      R_f[3,0] := -0.22841774;
      R_f[3,1] := 0.40559068;
      R_f[3,2] := 0.57486951;
      R_f[3,3] := 2.06207776;
      R_f[3,4] := -0.55732775;
      R_f[3,5] := 0.09659977;
      R_f[3,6] := -0.42354828;
      R_f[3,7] := -0.45963588;
      R_f[3,8] := -0.44553128;
      R_f[3,9] := -0.58046556;
      R_f[3,10] := -0.80908269;
      R_f[3,11] := -0.36142787;
      R_f[3,12] := 0.31985673;
      R_f[3,13] := -0.12466143;
      R_f[3,14] := 0.03553643;
      R_f[3,15] := -0.42549297;
      R_f[3,16] := -0.98859489;
      R_f[3,17] := 0.11508524;
      R_f[3,18] := 0.12030809;
      R_f[3,19] := 0.61023998;
      R_f[3,20] := -0.23926187;
      R_f[3,21] := -0.02740595;
      R_f[3,22] := 0.06562693;
      R_f[3,23] := 0.00750753;
      R_f[3,24] := 0.04459137;
      R_f[3,25] := 0.22271563;
      R_f[3,26] := -0.04020920;
      R_f[3,27] := 0.33254516;
      R_f[3,28] := 0.11126116;
      R_f[3,29] := -0.20861124;
      R_f[3,30] := 0.21898773;
      R_f[3,31] := 0.09003633;
      R_f[4,0] := -0.29503077;
      R_f[4,1] := 0.29277351;
      R_f[4,2] := -0.33615652;
      R_f[4,3] := 0.01891872;
      R_f[4,4] := -1.01232004;
      R_f[4,5] := 0.50957382;
      R_f[4,6] := -0.09908187;
      R_f[4,7] := -0.13480274;
      R_f[4,8] := -0.03347661;
      R_f[4,9] := 0.26127309;
      R_f[4,10] := -0.11804081;
      R_f[4,11] := -0.43345410;
      R_f[4,12] := 0.43429026;
      R_f[4,13] := -0.29253858;
      R_f[4,14] := 0.34731063;
      R_f[4,15] := -0.31193343;
      R_f[4,16] := 0.44109902;
      R_f[4,17] := 0.05499700;
      R_f[4,18] := -0.03124390;
      R_f[4,19] := -0.06733673;
      R_f[4,20] := 0.53314525;
      R_f[4,21] := 0.02740945;
      R_f[4,22] := -0.01510098;
      R_f[4,23] := 0.22094952;
      R_f[4,24] := -0.13394623;
      R_f[4,25] := 0.16025461;
      R_f[4,26] := 0.41375709;
      R_f[4,27] := -0.68666464;
      R_f[4,28] := 0.17169803;
      R_f[4,29] := -0.06553656;
      R_f[4,30] := -0.27536944;
      R_f[4,31] := 0.20692281;
      R_f[5,0] := 0.33732611;
      R_f[5,1] := 0.40928459;
      R_f[5,2] := -0.75300062;
      R_f[5,3] := -0.55881333;
      R_f[5,4] := 0.83829790;
      R_f[5,5] := -1.23661423;
      R_f[5,6] := -0.00860018;
      R_f[5,7] := 0.15366301;
      R_f[5,8] := 0.83814925;
      R_f[5,9] := -0.83846211;
      R_f[5,10] := 0.15663271;
      R_f[5,11] := -0.53920645;
      R_f[5,12] := -0.22816044;
      R_f[5,13] := -0.81048518;
      R_f[5,14] := 0.00169420;
      R_f[5,15] := 0.16230814;
      R_f[5,16] := 0.78781903;
      R_f[5,17] := -0.45289493;
      R_f[5,18] := 0.47988066;
      R_f[5,19] := -0.27889726;
      R_f[5,20] := 0.08924929;
      R_f[5,21] := -0.53515106;
      R_f[5,22] := 0.83308595;
      R_f[5,23] := 0.17609777;
      R_f[5,24] := -0.01040109;
      R_f[5,25] := 0.30510819;
      R_f[5,26] := 0.55807745;
      R_f[5,27] := 0.10998377;
      R_f[5,28] := -0.16242138;
      R_f[5,29] := -0.67912698;
      R_f[5,30] := -0.18073113;
      R_f[5,31] := 0.44595328;
      R_f[6,0] := -0.02960970;
      R_f[6,1] := 0.14120346;
      R_f[6,2] := -0.19232050;
      R_f[6,3] := -0.20220532;
      R_f[6,4] := 0.59759414;
      R_f[6,5] := 0.07536479;
      R_f[6,6] := 0.45140901;
      R_f[6,7] := -0.13872539;
      R_f[6,8] := 0.89296800;
      R_f[6,9] := -0.13736337;
      R_f[6,10] := 0.20182616;
      R_f[6,11] := -0.13915065;
      R_f[6,12] := -0.17636664;
      R_f[6,13] := -0.37117252;
      R_f[6,14] := 0.26237535;
      R_f[6,15] := -0.13584390;
      R_f[6,16] := 0.23492494;
      R_f[6,17] := -0.51170081;
      R_f[6,18] := -0.13849613;
      R_f[6,19] := -0.06773239;
      R_f[6,20] := 0.28203338;
      R_f[6,21] := 0.02628134;
      R_f[6,22] := 0.24086651;
      R_f[6,23] := 0.14421909;
      R_f[6,24] := 0.81928957;
      R_f[6,25] := 0.33552960;
      R_f[6,26] := -0.28975615;
      R_f[6,27] := 0.02547251;
      R_f[6,28] := 0.20271114;
      R_f[6,29] := -0.14385954;
      R_f[6,30] := 0.29766709;
      R_f[6,31] := -0.40624860;
      R_f[7,0] := 0.61828715;
      R_f[7,1] := 0.51957172;
      R_f[7,2] := 0.07738917;
      R_f[7,3] := -0.00875778;
      R_f[7,4] := 0.67404419;
      R_f[7,5] := 0.11073278;
      R_f[7,6] := -0.37006202;
      R_f[7,7] := 1.03556788;
      R_f[7,8] := 0.70712101;
      R_f[7,9] := -0.56803280;
      R_f[7,10] := -0.06974930;
      R_f[7,11] := 0.14248914;
      R_f[7,12] := 0.66664493;
      R_f[7,13] := -0.50647444;
      R_f[7,14] := 0.28662270;
      R_f[7,15] := 0.16329370;
      R_f[7,16] := -0.00441234;
      R_f[7,17] := -0.22685143;
      R_f[7,18] := -0.64886677;
      R_f[7,19] := -0.03913877;
      R_f[7,20] := 0.57906586;
      R_f[7,21] := 0.41091961;
      R_f[7,22] := 0.19402935;
      R_f[7,23] := -0.56783932;
      R_f[7,24] := 0.59809852;
      R_f[7,25] := 0.22131553;
      R_f[7,26] := 0.01115896;
      R_f[7,27] := 0.20468640;
      R_f[7,28] := -0.69074368;
      R_f[7,29] := -0.22870129;
      R_f[7,30] := 0.38742521;
      R_f[7,31] := -0.17464639;
      R_f[8,0] := -0.01413119;
      R_f[8,1] := -0.01563436;
      R_f[8,2] := 0.04907341;
      R_f[8,3] := 0.13082743;
      R_f[8,4] := -0.14134008;
      R_f[8,5] := -0.09485538;
      R_f[8,6] := -0.31782639;
      R_f[8,7] := -0.00754579;
      R_f[8,8] := -0.68271863;
      R_f[8,9] := 0.43590066;
      R_f[8,10] := -0.16523221;
      R_f[8,11] := 0.20073125;
      R_f[8,12] := -0.47652704;
      R_f[8,13] := 0.18128465;
      R_f[8,14] := -0.62839359;
      R_f[8,15] := -0.25646719;
      R_f[8,16] := -0.23885600;
      R_f[8,17] := 0.13142671;
      R_f[8,18] := 0.48771819;
      R_f[8,19] := -0.49085858;
      R_f[8,20] := -0.18839863;
      R_f[8,21] := -0.43685639;
      R_f[8,22] := 0.02705371;
      R_f[8,23] := -0.05543226;
      R_f[8,24] := -0.38585073;
      R_f[8,25] := 0.06531966;
      R_f[8,26] := -0.15446883;
      R_f[8,27] := 0.05854914;
      R_f[8,28] := -0.30904549;
      R_f[8,29] := 0.05056802;
      R_f[8,30] := -0.41357008;
      R_f[8,31] := 0.20621774;
      R_f[9,0] := -0.83740795;
      R_f[9,1] := -0.06988145;
      R_f[9,2] := -0.01356161;
      R_f[9,3] := 0.08127308;
      R_f[9,4] := -0.45402661;
      R_f[9,5] := 0.38458407;
      R_f[9,6] := 0.26937473;
      R_f[9,7] := -0.32646099;
      R_f[9,8] := -0.91716331;
      R_f[9,9] := 1.38183928;
      R_f[9,10] := 0.15634774;
      R_f[9,11] := -0.17276365;
      R_f[9,12] := -0.16843350;
      R_f[9,13] := -0.24043344;
      R_f[9,14] := -1.08728600;
      R_f[9,15] := -0.43865058;
      R_f[9,16] := 0.03624129;
      R_f[9,17] := 0.46195465;
      R_f[9,18] := 0.28181869;
      R_f[9,19] := 0.00515404;
      R_f[9,20] := -0.05451173;
      R_f[9,21] := 0.29636249;
      R_f[9,22] := -0.61817378;
      R_f[9,23] := 0.29860359;
      R_f[9,24] := -0.34871268;
      R_f[9,25] := 0.11697577;
      R_f[9,26] := 0.78417259;
      R_f[9,27] := 0.71926928;
      R_f[9,28] := -0.20325977;
      R_f[9,29] := 0.14632353;
      R_f[9,30] := -0.25228071;
      R_f[9,31] := -0.32943490;
      R_f[10,0] := 0.38591698;
      R_f[10,1] := 0.00522286;
      R_f[10,2] := -0.48348549;
      R_f[10,3] := 0.96521038;
      R_f[10,4] := -0.32313466;
      R_f[10,5] := 0.30804583;
      R_f[10,6] := -0.79955953;
      R_f[10,7] := -0.31883714;
      R_f[10,8] := -0.90835553;
      R_f[10,9] := 0.30884159;
      R_f[10,10] := -1.16350293;
      R_f[10,11] := -0.63253200;
      R_f[10,12] := 0.59796506;
      R_f[10,13] := 0.48238036;
      R_f[10,14] := -0.10394208;
      R_f[10,15] := 0.16137904;
      R_f[10,16] := 0.11384938;
      R_f[10,17] := 1.00142598;
      R_f[10,18] := -0.75928485;
      R_f[10,19] := 0.28338146;
      R_f[10,20] := -0.95777762;
      R_f[10,21] := -0.61350137;
      R_f[10,22] := -0.70301116;
      R_f[10,23] := 0.22109440;
      R_f[10,24] := 0.32511491;
      R_f[10,25] := 0.58860904;
      R_f[10,26] := -0.02545941;
      R_f[10,27] := 0.26207218;
      R_f[10,28] := 0.75892609;
      R_f[10,29] := -0.47240314;
      R_f[10,30] := 0.02046607;
      R_f[10,31] := -0.29343525;
      R_f[11,0] := 0.63524234;
      R_f[11,1] := 0.13768600;
      R_f[11,2] := -0.28915507;
      R_f[11,3] := -0.18023908;
      R_f[11,4] := -0.26212382;
      R_f[11,5] := -0.55292249;
      R_f[11,6] := 0.16202901;
      R_f[11,7] := 0.35055608;
      R_f[11,8] := 0.59746683;
      R_f[11,9] := -0.60563761;
      R_f[11,10] := -0.04891396;
      R_f[11,11] := 1.17771423;
      R_f[11,12] := -0.31640816;
      R_f[11,13] := -0.11039021;
      R_f[11,14] := -0.08756445;
      R_f[11,15] := 0.00601315;
      R_f[11,16] := 0.32191852;
      R_f[11,17] := -0.90107346;
      R_f[11,18] := -0.47469705;
      R_f[11,19] := 0.05416169;
      R_f[11,20] := -0.09831773;
      R_f[11,21] := 0.10362659;
      R_f[11,22] := -0.00615723;
      R_f[11,23] := -0.13419445;
      R_f[11,24] := 0.07473942;
      R_f[11,25] := 0.45523170;
      R_f[11,26] := 0.17231539;
      R_f[11,27] := 0.18330109;
      R_f[11,28] := -0.33154044;
      R_f[11,29] := 0.00715767;
      R_f[11,30] := 0.02798121;
      R_f[11,31] := 0.12936890;
      R_f[12,0] := 0.52463913;
      R_f[12,1] := 1.23480833;
      R_f[12,2] := -0.26183358;
      R_f[12,3] := 0.29687256;
      R_f[12,4] := 0.12944640;
      R_f[12,5] := -0.64208639;
      R_f[12,6] := 0.14092363;
      R_f[12,7] := 0.29900426;
      R_f[12,8] := -0.38989353;
      R_f[12,9] := -0.15832269;
      R_f[12,10] := 0.38569406;
      R_f[12,11] := -0.49528036;
      R_f[12,12] := 0.83373916;
      R_f[12,13] := -0.42694458;
      R_f[12,14] := 0.76566309;
      R_f[12,15] := -0.48013216;
      R_f[12,16] := 0.40656197;
      R_f[12,17] := -0.31445476;
      R_f[12,18] := 0.24111255;
      R_f[12,19] := -0.19961938;
      R_f[12,20] := -0.11154682;
      R_f[12,21] := 0.33029765;
      R_f[12,22] := -0.13147451;
      R_f[12,23] := -0.03679356;
      R_f[12,24] := 0.17805246;
      R_f[12,25] := 0.05382822;
      R_f[12,26] := 0.43463483;
      R_f[12,27] := 0.27920336;
      R_f[12,28] := 0.55672109;
      R_f[12,29] := -0.69647855;
      R_f[12,30] := 0.65581310;
      R_f[12,31] := 0.12511645;
      R_f[13,0] := 0.23202457;
      R_f[13,1] := 0.62695414;
      R_f[13,2] := -0.71075511;
      R_f[13,3] := -0.91361868;
      R_f[13,4] := 1.39223123;
      R_f[13,5] := 0.40526325;
      R_f[13,6] := 0.07239435;
      R_f[13,7] := 0.16743791;
      R_f[13,8] := 0.89612418;
      R_f[13,9] := -0.92080438;
      R_f[13,10] := 0.23565021;
      R_f[13,11] := 0.41098762;
      R_f[13,12] := -0.37411463;
      R_f[13,13] := -0.37083071;
      R_f[13,14] := 0.21330817;
      R_f[13,15] := 0.32418102;
      R_f[13,16] := 0.64384466;
      R_f[13,17] := -0.70755357;
      R_f[13,18] := -0.60732776;
      R_f[13,19] := -0.31852406;
      R_f[13,20] := 0.38003522;
      R_f[13,21] := -0.38526192;
      R_f[13,22] := 0.85999751;
      R_f[13,23] := 0.08276569;
      R_f[13,24] := 0.52139038;
      R_f[13,25] := -0.09750945;
      R_f[13,26] := -0.19196609;
      R_f[13,27] := -0.18892166;
      R_f[13,28] := 0.12520945;
      R_f[13,29] := -0.40455785;
      R_f[13,30] := 0.87176305;
      R_f[13,31] := -0.29801390;
      R_f[14,0] := 0.08073674;
      R_f[14,1] := -0.22958316;
      R_f[14,2] := 0.39506468;
      R_f[14,3] := -0.29865783;
      R_f[14,4] := -0.24071212;
      R_f[14,5] := -0.54502225;
      R_f[14,6] := -0.22081053;
      R_f[14,7] := 0.11199540;
      R_f[14,8] := 0.39893955;
      R_f[14,9] := -0.00592328;
      R_f[14,10] := -0.56832987;
      R_f[14,11] := 0.19659449;
      R_f[14,12] := 0.57248878;
      R_f[14,13] := 0.22812998;
      R_f[14,14] := -0.08929932;
      R_f[14,15] := -0.43194354;
      R_f[14,16] := 0.15896702;
      R_f[14,17] := -0.12431962;
      R_f[14,18] := 0.43860698;
      R_f[14,19] := -0.23576687;
      R_f[14,20] := 0.12837251;
      R_f[14,21] := -0.08831814;
      R_f[14,22] := -0.12136080;
      R_f[14,23] := 0.56518930;
      R_f[14,24] := -0.46596053;
      R_f[14,25] := 0.19473872;
      R_f[14,26] := 0.19937690;
      R_f[14,27] := -1.21616924;
      R_f[14,28] := 0.46861416;
      R_f[14,29] := -0.24986319;
      R_f[14,30] := -0.61549062;
      R_f[14,31] := 0.33290240;
      R_f[15,0] := 0.31359208;
      R_f[15,1] := 0.33051741;
      R_f[15,2] := 0.15030840;
      R_f[15,3] := -0.38865900;
      R_f[15,4] := 0.06516448;
      R_f[15,5] := -0.32763284;
      R_f[15,6] := 0.21778707;
      R_f[15,7] := 0.23249651;
      R_f[15,8] := 0.02938646;
      R_f[15,9] := 0.06135718;
      R_f[15,10] := -0.27028698;
      R_f[15,11] := 0.40001541;
      R_f[15,12] := -0.00793086;
      R_f[15,13] := 0.00380884;
      R_f[15,14] := 0.08370329;
      R_f[15,15] := -0.22548552;
      R_f[15,16] := 0.02933858;
      R_f[15,17] := -0.35302344;
      R_f[15,18] := -0.25063863;
      R_f[15,19] := 0.28370765;
      R_f[15,20] := 0.04397562;
      R_f[15,21] := -0.07230925;
      R_f[15,22] := -0.09505362;
      R_f[15,23] := 0.15444055;
      R_f[15,24] := -0.02045420;
      R_f[15,25] := -0.14273162;
      R_f[15,26] := 0.37428376;
      R_f[15,27] := -0.05992498;
      R_f[15,28] := 0.16830987;
      R_f[15,29] := -0.32088986;
      R_f[15,30] := -0.33436120;
      R_f[15,31] := -0.37953538;
      R_f[16,0] := -0.26587957;
      R_f[16,1] := -0.31207001;
      R_f[16,2] := 0.50653142;
      R_f[16,3] := 1.14224505;
      R_f[16,4] := -0.61703724;
      R_f[16,5] := 0.13980502;
      R_f[16,6] := -0.14207593;
      R_f[16,7] := 0.39799580;
      R_f[16,8] := -0.42795599;
      R_f[16,9] := 0.49218190;
      R_f[16,10] := -0.02379325;
      R_f[16,11] := -0.01251386;
      R_f[16,12] := 0.81707931;
      R_f[16,13] := 0.56178325;
      R_f[16,14] := -0.41181156;
      R_f[16,15] := -0.34066352;
      R_f[16,16] := -0.47481647;
      R_f[16,17] := 0.51806176;
      R_f[16,18] := 0.20107090;
      R_f[16,19] := 0.04892090;
      R_f[16,20] := -0.22273828;
      R_f[16,21] := 0.42268997;
      R_f[16,22] := -0.21690965;
      R_f[16,23] := 0.55266404;
      R_f[16,24] := -0.78800714;
      R_f[16,25] := -0.40029246;
      R_f[16,26] := 0.31856278;
      R_f[16,27] := 0.15422256;
      R_f[16,28] := 0.08612204;
      R_f[16,29] := 0.27195919;
      R_f[16,30] := -0.04387485;
      R_f[16,31] := -0.06196566;
      R_f[17,0] := 0.05910539;
      R_f[17,1] := -0.21845020;
      R_f[17,2] := -0.64325720;
      R_f[17,3] := -0.17311564;
      R_f[17,4] := -0.05836086;
      R_f[17,5] := 0.08543847;
      R_f[17,6] := 0.43946153;
      R_f[17,7] := 0.30724356;
      R_f[17,8] := 0.06860433;
      R_f[17,9] := 0.62805259;
      R_f[17,10] := 0.54351902;
      R_f[17,11] := 0.07233211;
      R_f[17,12] := -0.29924318;
      R_f[17,13] := -0.46094373;
      R_f[17,14] := -0.06874729;
      R_f[17,15] := 0.24842280;
      R_f[17,16] := -0.51377529;
      R_f[17,17] := 1.53367448;
      R_f[17,18] := 0.33991754;
      R_f[17,19] := 0.21408086;
      R_f[17,20] := -0.02237522;
      R_f[17,21] := -0.02311720;
      R_f[17,22] := 0.23792864;
      R_f[17,23] := 0.21117508;
      R_f[17,24] := -0.01755552;
      R_f[17,25] := -0.14541535;
      R_f[17,26] := 0.62708884;
      R_f[17,27] := 0.03084901;
      R_f[17,28] := -0.38820636;
      R_f[17,29] := -0.19554625;
      R_f[17,30] := 0.06806003;
      R_f[17,31] := -0.30774286;
      R_f[18,0] := 0.16866495;
      R_f[18,1] := 0.42400992;
      R_f[18,2] := -0.36475778;
      R_f[18,3] := -0.46353397;
      R_f[18,4] := -0.23605427;
      R_f[18,5] := -0.39058918;
      R_f[18,6] := 0.24388304;
      R_f[18,7] := -0.24780002;
      R_f[18,8] := -0.12100184;
      R_f[18,9] := -0.35586256;
      R_f[18,10] := 0.54968441;
      R_f[18,11] := -0.25823474;
      R_f[18,12] := -0.37975135;
      R_f[18,13] := 0.10739443;
      R_f[18,14] := 0.02995439;
      R_f[18,15] := 0.37767676;
      R_f[18,16] := -0.06366078;
      R_f[18,17] := 0.32446918;
      R_f[18,18] := 0.87205279;
      R_f[18,19] := -0.05647478;
      R_f[18,20] := -0.19952400;
      R_f[18,21] := -0.61423117;
      R_f[18,22] := 0.49618649;
      R_f[18,23] := -0.15967572;
      R_f[18,24] := 0.65420824;
      R_f[18,25] := 0.12151071;
      R_f[18,26] := 0.31860438;
      R_f[18,27] := 0.02739185;
      R_f[18,28] := -0.66384917;
      R_f[18,29] := 0.17025499;
      R_f[18,30] := -0.25605354;
      R_f[18,31] := 0.52890509;
      R_f[19,0] := 0.65365380;
      R_f[19,1] := 0.10235491;
      R_f[19,2] := 0.62065804;
      R_f[19,3] := 0.10225008;
      R_f[19,4] := -0.45779619;
      R_f[19,5] := -0.42509148;
      R_f[19,6] := -0.48240736;
      R_f[19,7] := -0.41890648;
      R_f[19,8] := 0.51948655;
      R_f[19,9] := 0.22051780;
      R_f[19,10] := -0.32477748;
      R_f[19,11] := -1.20024562;
      R_f[19,12] := 0.22928596;
      R_f[19,13] := 0.10820945;
      R_f[19,14] := -0.23491700;
      R_f[19,15] := -0.34898815;
      R_f[19,16] := -0.93565780;
      R_f[19,17] := 0.20988458;
      R_f[19,18] := -0.31584072;
      R_f[19,19] := -0.02921623;
      R_f[19,20] := -0.26133105;
      R_f[19,21] := 0.63414830;
      R_f[19,22] := -0.26187015;
      R_f[19,23] := 0.26986319;
      R_f[19,24] := -0.16388878;
      R_f[19,25] := 0.39682811;
      R_f[19,26] := 0.23186836;
      R_f[19,27] := 0.33898479;
      R_f[19,28] := -0.19298120;
      R_f[19,29] := 0.05988296;
      R_f[19,30] := 0.30527696;
      R_f[19,31] := 0.35504943;
      R_f[20,0] := 0.60740626;
      R_f[20,1] := 0.68342733;
      R_f[20,2] := -0.56973433;
      R_f[20,3] := 0.30702043;
      R_f[20,4] := 0.63084090;
      R_f[20,5] := -0.76327389;
      R_f[20,6] := -0.16775738;
      R_f[20,7] := 0.29119602;
      R_f[20,8] := -0.24701932;
      R_f[20,9] := -0.93371648;
      R_f[20,10] := 0.65781426;
      R_f[20,11] := -0.03017730;
      R_f[20,12] := -0.59253180;
      R_f[20,13] := -1.06371450;
      R_f[20,14] := 0.88938069;
      R_f[20,15] := 0.20159939;
      R_f[20,16] := 0.31710625;
      R_f[20,17] := 0.17246717;
      R_f[20,18] := 0.76323175;
      R_f[20,19] := 0.10229112;
      R_f[20,20] := -0.21142122;
      R_f[20,21] := -0.31407952;
      R_f[20,22] := -0.34694698;
      R_f[20,23] := -0.14305308;
      R_f[20,24] := 0.66643405;
      R_f[20,25] := -0.32228628;
      R_f[20,26] := 0.18264067;
      R_f[20,27] := 0.21311571;
      R_f[20,28] := 0.15977044;
      R_f[20,29] := 0.35266665;
      R_f[20,30] := 0.07271075;
      R_f[20,31] := 0.90672767;
      R_f[21,0] := 0.63794458;
      R_f[21,1] := -0.07306197;
      R_f[21,2] := -0.33461115;
      R_f[21,3] := 0.07822674;
      R_f[21,4] := 0.38671464;
      R_f[21,5] := -0.92790735;
      R_f[21,6] := -0.12789188;
      R_f[21,7] := -0.12363939;
      R_f[21,8] := 0.18649052;
      R_f[21,9] := -0.47208816;
      R_f[21,10] := -0.51584691;
      R_f[21,11] := 0.18042590;
      R_f[21,12] := 0.45089826;
      R_f[21,13] := 0.13358073;
      R_f[21,14] := 0.68462294;
      R_f[21,15] := -0.50330412;
      R_f[21,16] := -0.00928727;
      R_f[21,17] := -0.18551630;
      R_f[21,18] := 0.23045629;
      R_f[21,19] := -0.24903311;
      R_f[21,20] := -0.21607880;
      R_f[21,21] := 1.09473407;
      R_f[21,22] := 0.22049566;
      R_f[21,23] := 0.00980196;
      R_f[21,24] := 0.42017451;
      R_f[21,25] := 0.18463401;
      R_f[21,26] := 0.72073048;
      R_f[21,27] := 0.08499105;
      R_f[21,28] := -0.05317052;
      R_f[21,29] := 0.01483204;
      R_f[21,30] := 0.42573896;
      R_f[21,31] := 0.58880693;
      R_f[22,0] := 0.52571583;
      R_f[22,1] := 0.74352360;
      R_f[22,2] := -0.42845920;
      R_f[22,3] := -0.12134498;
      R_f[22,4] := -0.33517385;
      R_f[22,5] := -0.53988433;
      R_f[22,6] := -0.19025023;
      R_f[22,7] := -0.33218449;
      R_f[22,8] := -0.56198525;
      R_f[22,9] := 0.06062734;
      R_f[22,10] := -0.15277702;
      R_f[22,11] := -0.15610690;
      R_f[22,12] := -0.85074830;
      R_f[22,13] := -0.27995047;
      R_f[22,14] := 0.04608161;
      R_f[22,15] := 0.20265953;
      R_f[22,16] := 0.61842918;
      R_f[22,17] := -0.35963365;
      R_f[22,18] := 0.32028535;
      R_f[22,19] := 0.40971312;
      R_f[22,20] := 0.07105415;
      R_f[22,21] := -0.26550075;
      R_f[22,22] := 0.32755789;
      R_f[22,23] := -0.53670889;
      R_f[22,24] := 0.81352252;
      R_f[22,25] := 0.17814557;
      R_f[22,26] := -0.27500603;
      R_f[22,27] := 0.17979041;
      R_f[22,28] := 0.77811944;
      R_f[22,29] := -0.40859875;
      R_f[22,30] := -0.01199397;
      R_f[22,31] := 0.16662607;
      R_f[23,0] := 0.18513951;
      R_f[23,1] := -0.36498722;
      R_f[23,2] := 0.12142582;
      R_f[23,3] := 0.06119955;
      R_f[23,4] := 0.18143424;
      R_f[23,5] := -0.15825206;
      R_f[23,6] := -0.56776536;
      R_f[23,7] := 0.03979553;
      R_f[23,8] := -0.57782358;
      R_f[23,9] := 0.17007102;
      R_f[23,10] := 0.03401264;
      R_f[23,11] := 0.30232838;
      R_f[23,12] := 0.60225219;
      R_f[23,13] := 0.13679615;
      R_f[23,14] := -0.17490226;
      R_f[23,15] := -0.38221130;
      R_f[23,16] := -0.35548767;
      R_f[23,17] := -0.11720476;
      R_f[23,18] := 0.10709175;
      R_f[23,19] := 0.27031457;
      R_f[23,20] := -0.21203364;
      R_f[23,21] := 0.10817976;
      R_f[23,22] := -0.02741619;
      R_f[23,23] := -0.12317895;
      R_f[23,24] := -0.43592772;
      R_f[23,25] := -0.06452787;
      R_f[23,26] := 0.23145935;
      R_f[23,27] := -0.13228178;
      R_f[23,28] := -0.27505627;
      R_f[23,29] := 0.07636941;
      R_f[23,30] := -0.40810692;
      R_f[23,31] := 0.42898092;
      R_f[24,0] := 0.28041553;
      R_f[24,1] := 0.35192281;
      R_f[24,2] := -0.45653370;
      R_f[24,3] := -0.39068758;
      R_f[24,4] := 0.59820068;
      R_f[24,5] := -0.14331487;
      R_f[24,6] := -0.16312519;
      R_f[24,7] := 0.20082375;
      R_f[24,8] := 0.85522902;
      R_f[24,9] := -1.29532707;
      R_f[24,10] := 0.44740444;
      R_f[24,11] := -0.42685062;
      R_f[24,12] := -0.38446230;
      R_f[24,13] := -0.25391304;
      R_f[24,14] := 0.57489002;
      R_f[24,15] := -0.11480054;
      R_f[24,16] := 0.49371004;
      R_f[24,17] := -0.34504244;
      R_f[24,18] := 0.08720941;
      R_f[24,19] := -0.72877926;
      R_f[24,20] := -0.04864010;
      R_f[24,21] := -0.53587073;
      R_f[24,22] := 0.82679683;
      R_f[24,23] := -0.64950413;
      R_f[24,24] := 0.71601194;
      R_f[24,25] := 0.38295448;
      R_f[24,26] := 0.40242442;
      R_f[24,27] := 0.20521010;
      R_f[24,28] := -0.03906753;
      R_f[24,29] := -0.60810322;
      R_f[24,30] := 0.03209632;
      R_f[24,31] := -0.01952329;
      R_f[25,0] := 0.24457985;
      R_f[25,1] := -1.02144086;
      R_f[25,2] := -1.15114701;
      R_f[25,3] := -0.35912865;
      R_f[25,4] := 0.10526828;
      R_f[25,5] := -0.20179662;
      R_f[25,6] := -0.08682156;
      R_f[25,7] := -0.53071922;
      R_f[25,8] := 0.78854895;
      R_f[25,9] := -0.39259291;
      R_f[25,10] := 0.01843655;
      R_f[25,11] := -0.56601465;
      R_f[25,12] := -0.02357278;
      R_f[25,13] := -0.37074372;
      R_f[25,14] := -0.04764435;
      R_f[25,15] := 0.07631879;
      R_f[25,16] := 0.14908385;
      R_f[25,17] := -0.22848843;
      R_f[25,18] := 0.07038445;
      R_f[25,19] := -0.21256164;
      R_f[25,20] := -0.51917696;
      R_f[25,21] := -0.13761941;
      R_f[25,22] := 1.10180664;
      R_f[25,23] := -0.01601213;
      R_f[25,24] := 0.33799487;
      R_f[25,25] := 0.74898493;
      R_f[25,26] := 0.10358041;
      R_f[25,27] := -0.17927809;
      R_f[25,28] := -0.14816135;
      R_f[25,29] := -0.15051788;
      R_f[25,30] := 0.32431662;
      R_f[25,31] := -0.06228854;
      R_f[26,0] := -0.17391884;
      R_f[26,1] := 0.40459314;
      R_f[26,2] := 0.23582034;
      R_f[26,3] := 0.27855241;
      R_f[26,4] := 0.41587636;
      R_f[26,5] := -0.06871118;
      R_f[26,6] := -0.18198022;
      R_f[26,7] := 0.30424389;
      R_f[26,8] := 0.47402722;
      R_f[26,9] := 0.10770813;
      R_f[26,10] := 0.19400623;
      R_f[26,11] := 0.19763534;
      R_f[26,12] := 0.83919579;
      R_f[26,13] := -0.20429327;
      R_f[26,14] := 0.30284089;
      R_f[26,15] := -0.15002888;
      R_f[26,16] := 0.68186575;
      R_f[26,17] := 0.55425143;
      R_f[26,18] := 0.27912667;
      R_f[26,19] := 0.33006024;
      R_f[26,20] := 0.64902514;
      R_f[26,21] := -0.04681511;
      R_f[26,22] := 0.43274990;
      R_f[26,23] := -0.06403653;
      R_f[26,24] := 0.90166181;
      R_f[26,25] := -0.52762878;
      R_f[26,26] := -0.00969170;
      R_f[26,27] := -0.59007823;
      R_f[26,28] := 0.04513381;
      R_f[26,29] := -1.11053836;
      R_f[26,30] := -0.14078638;
      R_f[26,31] := 0.10301355;
      R_f[27,0] := 0.39776009;
      R_f[27,1] := 0.59193295;
      R_f[27,2] := -0.16674590;
      R_f[27,3] := -0.01398129;
      R_f[27,4] := 0.34197676;
      R_f[27,5] := -0.11277734;
      R_f[27,6] := -0.18087836;
      R_f[27,7] := -0.24809147;
      R_f[27,8] := 1.11544597;
      R_f[27,9] := -0.41635385;
      R_f[27,10] := 1.21610570;
      R_f[27,11] := -0.42330170;
      R_f[27,12] := -0.49244744;
      R_f[27,13] := -0.17151001;
      R_f[27,14] := -0.73654294;
      R_f[27,15] := 0.40863410;
      R_f[27,16] := 0.30207148;
      R_f[27,17] := -0.30706853;
      R_f[27,18] := 0.17934655;
      R_f[27,19] := -0.01947166;
      R_f[27,20] := 0.29237783;
      R_f[27,21] := -0.18835185;
      R_f[27,22] := -0.42462611;
      R_f[27,23] := -0.31352675;
      R_f[27,24] := 0.80565614;
      R_f[27,25] := 0.15593880;
      R_f[27,26] := -0.07164915;
      R_f[27,27] := 1.59558272;
      R_f[27,28] := -0.26499027;
      R_f[27,29] := -0.86730254;
      R_f[27,30] := 0.45258304;
      R_f[27,31] := -0.10650399;
      R_f[28,0] := 0.29013574;
      R_f[28,1] := 0.78875935;
      R_f[28,2] := -0.22047451;
      R_f[28,3] := 0.31630492;
      R_f[28,4] := 0.13784394;
      R_f[28,5] := -0.17747335;
      R_f[28,6] := -0.16462083;
      R_f[28,7] := 0.02444983;
      R_f[28,8] := 0.02157918;
      R_f[28,9] := -0.85899609;
      R_f[28,10] := 0.51003945;
      R_f[28,11] := 0.22153500;
      R_f[28,12] := -0.81957668;
      R_f[28,13] := 0.15229519;
      R_f[28,14] := -0.49981925;
      R_f[28,15] := -0.20841819;
      R_f[28,16] := 0.48134491;
      R_f[28,17] := -0.58209991;
      R_f[28,18] := -0.21895251;
      R_f[28,19] := -0.31777707;
      R_f[28,20] := 0.39952904;
      R_f[28,21] := 0.33487400;
      R_f[28,22] := 0.53231794;
      R_f[28,23] := 0.58753723;
      R_f[28,24] := 0.29652479;
      R_f[28,25] := 0.49816924;
      R_f[28,26] := -0.19129919;
      R_f[28,27] := 0.74723542;
      R_f[28,28] := 0.06283404;
      R_f[28,29] := -0.70639998;
      R_f[28,30] := 0.34521261;
      R_f[28,31] := -0.15957113;
      R_f[29,0] := 0.23835732;
      R_f[29,1] := -0.26068553;
      R_f[29,2] := -0.55099136;
      R_f[29,3] := -0.27018866;
      R_f[29,4] := -0.35758555;
      R_f[29,5] := 0.74466068;
      R_f[29,6] := 0.46339175;
      R_f[29,7] := -0.27842417;
      R_f[29,8] := 0.12199467;
      R_f[29,9] := -0.58916980;
      R_f[29,10] := 0.10298276;
      R_f[29,11] := -0.58598566;
      R_f[29,12] := 0.03986860;
      R_f[29,13] := 0.36140522;
      R_f[29,14] := 0.14722234;
      R_f[29,15] := -0.15363480;
      R_f[29,16] := 0.72394967;
      R_f[29,17] := -0.39522561;
      R_f[29,18] := -0.06369760;
      R_f[29,19] := -0.19733445;
      R_f[29,20] := -0.23108549;
      R_f[29,21] := 0.09581164;
      R_f[29,22] := 0.60348934;
      R_f[29,23] := 0.38583145;
      R_f[29,24] := -0.32982609;
      R_f[29,25] := 0.76995927;
      R_f[29,26] := 0.39173558;
      R_f[29,27] := -0.11436092;
      R_f[29,28] := -0.33975780;
      R_f[29,29] := -2.43963838;
      R_f[29,30] := 0.01613091;
      R_f[29,31] := 1.01884580;
      R_f[30,0] := 0.44902706;
      R_f[30,1] := -0.01531547;
      R_f[30,2] := 0.43428138;
      R_f[30,3] := 0.20990226;
      R_f[30,4] := 0.10665958;
      R_f[30,5] := -0.07787514;
      R_f[30,6] := -0.28534907;
      R_f[30,7] := -0.20589265;
      R_f[30,8] := -0.26249862;
      R_f[30,9] := 0.32755303;
      R_f[30,10] := 0.16526289;
      R_f[30,11] := 0.07607982;
      R_f[30,12] := 0.15522026;
      R_f[30,13] := 0.16349413;
      R_f[30,14] := -0.41222379;
      R_f[30,15] := -0.37317255;
      R_f[30,16] := -0.38004446;
      R_f[30,17] := -0.11156923;
      R_f[30,18] := -0.06939796;
      R_f[30,19] := 0.75725025;
      R_f[30,20] := 0.16113472;
      R_f[30,21] := 0.36386901;
      R_f[30,22] := 0.15552250;
      R_f[30,23] := -0.10594840;
      R_f[30,24] := -0.00384362;
      R_f[30,25] := -0.10023083;
      R_f[30,26] := 0.55560988;
      R_f[30,27] := 0.35110676;
      R_f[30,28] := -0.28105840;
      R_f[30,29] := -0.08273152;
      R_f[30,30] := 0.76468736;
      R_f[30,31] := 0.03726526;
      R_f[31,0] := 0.43319872;
      R_f[31,1] := 0.89265436;
      R_f[31,2] := -0.02175743;
      R_f[31,3] := -0.23646763;
      R_f[31,4] := -0.24073155;
      R_f[31,5] := -0.00261918;
      R_f[31,6] := -0.57301140;
      R_f[31,7] := -0.04121628;
      R_f[31,8] := -0.32528654;
      R_f[31,9] := -0.79124427;
      R_f[31,10] := -0.25563994;
      R_f[31,11] := 0.61876816;
      R_f[31,12] := -0.24966605;
      R_f[31,13] := -0.15887363;
      R_f[31,14] := -0.27610224;
      R_f[31,15] := -0.24292535;
      R_f[31,16] := -0.17999788;
      R_f[31,17] := -0.17289916;
      R_f[31,18] := 0.49396884;
      R_f[31,19] := 0.35957804;
      R_f[31,20] := -0.07121407;
      R_f[31,21] := 0.01738700;
      R_f[31,22] := 0.34174326;
      R_f[31,23] := -0.52943313;
      R_f[31,24] := -0.28900346;
      R_f[31,25] := 0.48076582;
      R_f[31,26] := -0.03657150;
      R_f[31,27] := 0.02927713;
      R_f[31,28] := -0.82611400;
      R_f[31,29] := -0.81384391;
      R_f[31,30] := -0.24894159;
      R_f[31,31] := 1.24944818;
      R_g[0,0] := -3.90892291;
      R_g[0,1] := -0.07594703;
      R_g[0,2] := -0.11032616;
      R_g[0,3] := -0.12472310;
      R_g[0,4] := -0.00621575;
      R_g[0,5] := 0.19935456;
      R_g[0,6] := -0.06362464;
      R_g[0,7] := -0.16034737;
      R_g[0,8] := 0.09810749;
      R_g[0,9] := 0.12010512;
      R_g[0,10] := 0.17773002;
      R_g[0,11] := -0.01798855;
      R_g[0,12] := -0.10235326;
      R_g[0,13] := 0.23832326;
      R_g[0,14] := 0.11828293;
      R_g[0,15] := -0.07939270;
      R_g[0,16] := -0.14808963;
      R_g[0,17] := 0.03173243;
      R_g[0,18] := 0.18550968;
      R_g[0,19] := -0.06182884;
      R_g[0,20] := 0.04494766;
      R_g[0,21] := -0.12930253;
      R_g[0,22] := -0.04077970;
      R_g[0,23] := 0.12853464;
      R_g[0,24] := 0.04193184;
      R_g[0,25] := 0.25337324;
      R_g[0,26] := -0.18417910;
      R_g[0,27] := -0.18281718;
      R_g[0,28] := 0.12372693;
      R_g[0,29] := 0.04042292;
      R_g[0,30] := -0.09040337;
      R_g[0,31] := 0.04066515;
      R_g[1,0] := 0.29689670;
      R_g[1,1] := -3.97663403;
      R_g[1,2] := 0.06429198;
      R_g[1,3] := 0.01962975;
      R_g[1,4] := -0.15935937;
      R_g[1,5] := 0.15787816;
      R_g[1,6] := 0.12121452;
      R_g[1,7] := 0.05212499;
      R_g[1,8] := 0.00120139;
      R_g[1,9] := -0.04333260;
      R_g[1,10] := -0.10989881;
      R_g[1,11] := 0.04567650;
      R_g[1,12] := -0.06217363;
      R_g[1,13] := 0.02787914;
      R_g[1,14] := -0.21347456;
      R_g[1,15] := 0.04342266;
      R_g[1,16] := 0.04235249;
      R_g[1,17] := -0.23068787;
      R_g[1,18] := 0.02733839;
      R_g[1,19] := 0.02264871;
      R_g[1,20] := -0.32929158;
      R_g[1,21] := -0.04880635;
      R_g[1,22] := -0.07773370;
      R_g[1,23] := -0.19768843;
      R_g[1,24] := 0.07725871;
      R_g[1,25] := -0.09810391;
      R_g[1,26] := 0.04568880;
      R_g[1,27] := 0.25973374;
      R_g[1,28] := -0.11771499;
      R_g[1,29] := 0.07775978;
      R_g[1,30] := 0.06788124;
      R_g[1,31] := -0.15774764;
      R_g[2,0] := 0.78595299;
      R_g[2,1] := -0.03254539;
      R_g[2,2] := -3.97857785;
      R_g[2,3] := 0.03195208;
      R_g[2,4] := -0.00134882;
      R_g[2,5] := 0.00648824;
      R_g[2,6] := 0.37531501;
      R_g[2,7] := 0.18654406;
      R_g[2,8] := 0.04044631;
      R_g[2,9] := 0.14008798;
      R_g[2,10] := -0.07232818;
      R_g[2,11] := 0.20235972;
      R_g[2,12] := -0.00854753;
      R_g[2,13] := -0.17538439;
      R_g[2,14] := 0.05945322;
      R_g[2,15] := -0.23242135;
      R_g[2,16] := 0.03825035;
      R_g[2,17] := 0.20309828;
      R_g[2,18] := -0.23156436;
      R_g[2,19] := 0.08224720;
      R_g[2,20] := -0.06343341;
      R_g[2,21] := -0.17136954;
      R_g[2,22] := 0.00879024;
      R_g[2,23] := -0.25821340;
      R_g[2,24] := 0.24464959;
      R_g[2,25] := -0.53886688;
      R_g[2,26] := -0.27455342;
      R_g[2,27] := -0.01048109;
      R_g[2,28] := -0.19415924;
      R_g[2,29] := -0.22414842;
      R_g[2,30] := -0.09919538;
      R_g[2,31] := -0.19051763;
      R_g[3,0] := -0.38880152;
      R_g[3,1] := 0.50711042;
      R_g[3,2] := 0.23847204;
      R_g[3,3] := -0.29851389;
      R_g[3,4] := 0.16963020;
      R_g[3,5] := 0.70479912;
      R_g[3,6] := -0.70167243;
      R_g[3,7] := -0.30499798;
      R_g[3,8] := 0.00119803;
      R_g[3,9] := 0.35383144;
      R_g[3,10] := -0.15565510;
      R_g[3,11] := 0.66530848;
      R_g[3,12] := 0.24109314;
      R_g[3,13] := 0.38931200;
      R_g[3,14] := 0.31814352;
      R_g[3,15] := -0.13152258;
      R_g[3,16] := 0.26083884;
      R_g[3,17] := 0.14622647;
      R_g[3,18] := 0.51298088;
      R_g[3,19] := 0.58923829;
      R_g[3,20] := 0.14318515;
      R_g[3,21] := 0.18607107;
      R_g[3,22] := -0.46340457;
      R_g[3,23] := -0.00351034;
      R_g[3,24] := -0.65315545;
      R_g[3,25] := 0.49816614;
      R_g[3,26] := -0.62532133;
      R_g[3,27] := -0.38666618;
      R_g[3,28] := 0.48155585;
      R_g[3,29] := -0.09343946;
      R_g[3,30] := -0.08817770;
      R_g[3,31] := 0.48095670;
      R_g[4,0] := -0.14076962;
      R_g[4,1] := 0.04399427;
      R_g[4,2] := -0.11605984;
      R_g[4,3] := -0.19373409;
      R_g[4,4] := -2.39188242;
      R_g[4,5] := 0.56221688;
      R_g[4,6] := -0.11971202;
      R_g[4,7] := -0.12293410;
      R_g[4,8] := 0.16898374;
      R_g[4,9] := 0.22141531;
      R_g[4,10] := 0.06616066;
      R_g[4,11] := 0.03161502;
      R_g[4,12] := 0.04760331;
      R_g[4,13] := -0.94796467;
      R_g[4,14] := -0.21785344;
      R_g[4,15] := 0.21287520;
      R_g[4,16] := -0.09627807;
      R_g[4,17] := 0.33276817;
      R_g[4,18] := 0.36361930;
      R_g[4,19] := 0.11621923;
      R_g[4,20] := 0.12379040;
      R_g[4,21] := 0.28268778;
      R_g[4,22] := 0.02451998;
      R_g[4,23] := 0.07576066;
      R_g[4,24] := 0.14458476;
      R_g[4,25] := -0.09326506;
      R_g[4,26] := -0.10546308;
      R_g[4,27] := 0.23316522;
      R_g[4,28] := -0.18263954;
      R_g[4,29] := 0.04596911;
      R_g[4,30] := 0.16661571;
      R_g[4,31] := -0.14460705;
      R_g[5,0] := 0.00607648;
      R_g[5,1] := -0.31199628;
      R_g[5,2] := -0.14311165;
      R_g[5,3] := -0.08406878;
      R_g[5,4] := -0.45707089;
      R_g[5,5] := -3.66744041;
      R_g[5,6] := -0.29590583;
      R_g[5,7] := -0.36582258;
      R_g[5,8] := -0.20673501;
      R_g[5,9] := 0.93654841;
      R_g[5,10] := 0.17411292;
      R_g[5,11] := -0.64996815;
      R_g[5,12] := -0.29004732;
      R_g[5,13] := -0.40815744;
      R_g[5,14] := -0.04872389;
      R_g[5,15] := 0.34239492;
      R_g[5,16] := -0.43735024;
      R_g[5,17] := 0.99700075;
      R_g[5,18] := 0.77893156;
      R_g[5,19] := 0.07795681;
      R_g[5,20] := -0.13708429;
      R_g[5,21] := -0.00024443;
      R_g[5,22] := 0.64380318;
      R_g[5,23] := 0.64613158;
      R_g[5,24] := 0.24253663;
      R_g[5,25] := 0.58237201;
      R_g[5,26] := 0.38992611;
      R_g[5,27] := -0.11605772;
      R_g[5,28] := 0.41215706;
      R_g[5,29] := 0.48312679;
      R_g[5,30] := -0.01841857;
      R_g[5,31] := 0.32900634;
      R_g[6,0] := 0.21044113;
      R_g[6,1] := 0.27635157;
      R_g[6,2] := 0.25911206;
      R_g[6,3] := 0.20687383;
      R_g[6,4] := 0.42254698;
      R_g[6,5] := -0.06129316;
      R_g[6,6] := -2.86810660;
      R_g[6,7] := 0.01530620;
      R_g[6,8] := 0.03624671;
      R_g[6,9] := -0.55880523;
      R_g[6,10] := -0.11955739;
      R_g[6,11] := 0.23940329;
      R_g[6,12] := 0.20675407;
      R_g[6,13] := 0.32029077;
      R_g[6,14] := -0.08033612;
      R_g[6,15] := 0.01886825;
      R_g[6,16] := 0.44635811;
      R_g[6,17] := -0.47127756;
      R_g[6,18] := -0.12253133;
      R_g[6,19] := -0.11386113;
      R_g[6,20] := 0.08486191;
      R_g[6,21] := -0.04622066;
      R_g[6,22] := 0.04315218;
      R_g[6,23] := -0.34449965;
      R_g[6,24] := 0.14451315;
      R_g[6,25] := -0.08523499;
      R_g[6,26] := -0.62968856;
      R_g[6,27] := -0.22461188;
      R_g[6,28] := -0.12706000;
      R_g[6,29] := -0.11077819;
      R_g[6,30] := 0.03170905;
      R_g[6,31] := 0.29694375;
      R_g[7,0] := -0.13013278;
      R_g[7,1] := -0.31679758;
      R_g[7,2] := -0.07822036;
      R_g[7,3] := 0.20828305;
      R_g[7,4] := -0.26236439;
      R_g[7,5] := -0.20191798;
      R_g[7,6] := -0.16079828;
      R_g[7,7] := -2.61546016;
      R_g[7,8] := -0.11710360;
      R_g[7,9] := 0.28043556;
      R_g[7,10] := 0.13310109;
      R_g[7,11] := 0.07384923;
      R_g[7,12] := -0.09096892;
      R_g[7,13] := -0.11528125;
      R_g[7,14] := -0.00921861;
      R_g[7,15] := -0.01645553;
      R_g[7,16] := 0.09885471;
      R_g[7,17] := 0.22595286;
      R_g[7,18] := 0.18649556;
      R_g[7,19] := 0.18633325;
      R_g[7,20] := -0.19093995;
      R_g[7,21] := -0.03887040;
      R_g[7,22] := -0.20446028;
      R_g[7,23] := 0.23285761;
      R_g[7,24] := -0.13019045;
      R_g[7,25] := 0.39875758;
      R_g[7,26] := 0.06689890;
      R_g[7,27] := 0.15852100;
      R_g[7,28] := 0.07758270;
      R_g[7,29] := 0.10765402;
      R_g[7,30] := 0.01027874;
      R_g[7,31] := 0.10162933;
      R_g[8,0] := 0.52049464;
      R_g[8,1] := -0.06498682;
      R_g[8,2] := 0.22293125;
      R_g[8,3] := -0.26280743;
      R_g[8,4] := 0.10941017;
      R_g[8,5] := 0.05232298;
      R_g[8,6] := 0.12105810;
      R_g[8,7] := -0.66948277;
      R_g[8,8] := -1.77637279;
      R_g[8,9] := 0.54212058;
      R_g[8,10] := 0.52014560;
      R_g[8,11] := 0.25420547;
      R_g[8,12] := -0.18584058;
      R_g[8,13] := -0.23701867;
      R_g[8,14] := -0.02562778;
      R_g[8,15] := -0.03259461;
      R_g[8,16] := 0.12165561;
      R_g[8,17] := -0.06605203;
      R_g[8,18] := 0.01967831;
      R_g[8,19] := 0.90615851;
      R_g[8,20] := -0.25498098;
      R_g[8,21] := -0.26732451;
      R_g[8,22] := -0.19817455;
      R_g[8,23] := 0.22149684;
      R_g[8,24] := 0.04186046;
      R_g[8,25] := 0.48240146;
      R_g[8,26] := 0.43705374;
      R_g[8,27] := 0.23106116;
      R_g[8,28] := 0.24622135;
      R_g[8,29] := -0.14498775;
      R_g[8,30] := 0.11009011;
      R_g[8,31] := 0.07813966;
      R_g[9,0] := 0.16880883;
      R_g[9,1] := -0.37774763;
      R_g[9,2] := 0.25193521;
      R_g[9,3] := 0.21604455;
      R_g[9,4] := -0.52223831;
      R_g[9,5] := -0.23418076;
      R_g[9,6] := 0.45371133;
      R_g[9,7] := 0.07293321;
      R_g[9,8] := -0.31331846;
      R_g[9,9] := -0.15017952;
      R_g[9,10] := 0.14813878;
      R_g[9,11] := -0.22082219;
      R_g[9,12] := 0.15378278;
      R_g[9,13] := 0.56576324;
      R_g[9,14] := -0.73613793;
      R_g[9,15] := 0.06151476;
      R_g[9,16] := 0.01810322;
      R_g[9,17] := 0.44917166;
      R_g[9,18] := -0.11428359;
      R_g[9,19] := -0.15660156;
      R_g[9,20] := 0.17290512;
      R_g[9,21] := 0.25610337;
      R_g[9,22] := -0.14287926;
      R_g[9,23] := 0.34086990;
      R_g[9,24] := 0.09738272;
      R_g[9,25] := -0.37799767;
      R_g[9,26] := -0.07600447;
      R_g[9,27] := 0.03889601;
      R_g[9,28] := 0.42590618;
      R_g[9,29] := 0.00751106;
      R_g[9,30] := 0.09643213;
      R_g[9,31] := -0.04677634;
      R_g[10,0] := 0.62866777;
      R_g[10,1] := 0.04863711;
      R_g[10,2] := -0.21369855;
      R_g[10,3] := -0.50630087;
      R_g[10,4] := 0.01089374;
      R_g[10,5] := -0.56738806;
      R_g[10,6] := 0.01197762;
      R_g[10,7] := -0.29552773;
      R_g[10,8] := -0.18157986;
      R_g[10,9] := 0.02497040;
      R_g[10,10] := -1.49921405;
      R_g[10,11] := 0.34377626;
      R_g[10,12] := -0.31496713;
      R_g[10,13] := 0.05581916;
      R_g[10,14] := 0.01296536;
      R_g[10,15] := 0.07040508;
      R_g[10,16] := -0.07418365;
      R_g[10,17] := -0.22070369;
      R_g[10,18] := 0.04132200;
      R_g[10,19] := 0.23620397;
      R_g[10,20] := -0.08386072;
      R_g[10,21] := -0.37729159;
      R_g[10,22] := 0.45501009;
      R_g[10,23] := -0.01450009;
      R_g[10,24] := -0.19233912;
      R_g[10,25] := 0.31541747;
      R_g[10,26] := -0.06635552;
      R_g[10,27] := 0.20700711;
      R_g[10,28] := 0.20695294;
      R_g[10,29] := -0.20757411;
      R_g[10,30] := -0.08001424;
      R_g[10,31] := -0.13325055;
      R_g[11,0] := -0.29314852;
      R_g[11,1] := -0.02125665;
      R_g[11,2] := -0.18892588;
      R_g[11,3] := -0.13230674;
      R_g[11,4] := -0.00237155;
      R_g[11,5] := 0.26988694;
      R_g[11,6] := -0.20133880;
      R_g[11,7] := -0.20377180;
      R_g[11,8] := 0.06723951;
      R_g[11,9] := 0.37048879;
      R_g[11,10] := -0.05555879;
      R_g[11,11] := -2.22307801;
      R_g[11,12] := 0.04293208;
      R_g[11,13] := -0.15140139;
      R_g[11,14] := 0.12092919;
      R_g[11,15] := 0.09615011;
      R_g[11,16] := -0.47221011;
      R_g[11,17] := 0.51846349;
      R_g[11,18] := 0.42216018;
      R_g[11,19] := -0.05934686;
      R_g[11,20] := -0.05716062;
      R_g[11,21] := -0.22358482;
      R_g[11,22] := -0.24511711;
      R_g[11,23] := 0.33101672;
      R_g[11,24] := -0.22553165;
      R_g[11,25] := 0.41420865;
      R_g[11,26] := 0.39840400;
      R_g[11,27] := -0.09501968;
      R_g[11,28] := 0.12650503;
      R_g[11,29] := -0.18914959;
      R_g[11,30] := 0.15498011;
      R_g[11,31] := 0.17820162;
      R_g[12,0] := -0.09561817;
      R_g[12,1] := -0.29961327;
      R_g[12,2] := -0.03527441;
      R_g[12,3] := -0.34987089;
      R_g[12,4] := -0.06521978;
      R_g[12,5] := 0.00181486;
      R_g[12,6] := -0.01615610;
      R_g[12,7] := -0.07030049;
      R_g[12,8] := 0.09657750;
      R_g[12,9] := 0.07639907;
      R_g[12,10] := 0.18752827;
      R_g[12,11] := 0.04013976;
      R_g[12,12] := -2.89481735;
      R_g[12,13] := 0.09838540;
      R_g[12,14] := -0.05623082;
      R_g[12,15] := 0.32070735;
      R_g[12,16] := -0.28874421;
      R_g[12,17] := -0.01434616;
      R_g[12,18] := 0.23362166;
      R_g[12,19] := 0.07646300;
      R_g[12,20] := 0.22999871;
      R_g[12,21] := -0.28788614;
      R_g[12,22] := -0.18580739;
      R_g[12,23] := -0.13602987;
      R_g[12,24] := -0.10257613;
      R_g[12,25] := 0.03445209;
      R_g[12,26] := -0.30460083;
      R_g[12,27] := 0.24534188;
      R_g[12,28] := -0.15457958;
      R_g[12,29] := 0.23796089;
      R_g[12,30] := 0.20219725;
      R_g[12,31] := -0.24078710;
      R_g[13,0] := 0.75326633;
      R_g[13,1] := 0.42503357;
      R_g[13,2] := 0.25508878;
      R_g[13,3] := 0.25160366;
      R_g[13,4] := 0.98365158;
      R_g[13,5] := -0.28989795;
      R_g[13,6] := 0.49180490;
      R_g[13,7] := 0.45266271;
      R_g[13,8] := -0.05704876;
      R_g[13,9] := -0.73466700;
      R_g[13,10] := -0.12915684;
      R_g[13,11] := 0.46727014;
      R_g[13,12] := 0.19765535;
      R_g[13,13] := -3.78172469;
      R_g[13,14] := -0.34034637;
      R_g[13,15] := -0.45915127;
      R_g[13,16] := 0.33600780;
      R_g[13,17] := -0.61412776;
      R_g[13,18] := -0.89968032;
      R_g[13,19] := 0.01249010;
      R_g[13,20] := -0.04839383;
      R_g[13,21] := -0.21840587;
      R_g[13,22] := -0.34433964;
      R_g[13,23] := -0.70232898;
      R_g[13,24] := 0.12399767;
      R_g[13,25] := -0.55529630;
      R_g[13,26] := -0.20899974;
      R_g[13,27] := 0.24549794;
      R_g[13,28] := -0.23520455;
      R_g[13,29] := -0.46935543;
      R_g[13,30] := -0.04612514;
      R_g[13,31] := -0.26909268;
      R_g[14,0] := -0.04362309;
      R_g[14,1] := -0.00786453;
      R_g[14,2] := 0.47990274;
      R_g[14,3] := -0.08678034;
      R_g[14,4] := 0.26148090;
      R_g[14,5] := -0.09519535;
      R_g[14,6] := 0.17877942;
      R_g[14,7] := -0.18717366;
      R_g[14,8] := 0.06691048;
      R_g[14,9] := 0.17936321;
      R_g[14,10] := 0.88007951;
      R_g[14,11] := -0.27552536;
      R_g[14,12] := 0.02279478;
      R_g[14,13] := -0.49624246;
      R_g[14,14] := -1.74626386;
      R_g[14,15] := 0.12173577;
      R_g[14,16] := -0.29647782;
      R_g[14,17] := 0.29125968;
      R_g[14,18] := 0.38394415;
      R_g[14,19] := 0.01893454;
      R_g[14,20] := -0.04434190;
      R_g[14,21] := -0.03771880;
      R_g[14,22] := -0.25166640;
      R_g[14,23] := -0.19271357;
      R_g[14,24] := 0.25045004;
      R_g[14,25] := -0.18070081;
      R_g[14,26] := 0.11899330;
      R_g[14,27] := -0.45145723;
      R_g[14,28] := -0.11598604;
      R_g[14,29] := 0.14603114;
      R_g[14,30] := 0.13819149;
      R_g[14,31] := -0.38187009;
      R_g[15,0] := 0.17263101;
      R_g[15,1] := 0.09476559;
      R_g[15,2] := 0.08820881;
      R_g[15,3] := 0.12526147;
      R_g[15,4] := 0.06413334;
      R_g[15,5] := -0.39505017;
      R_g[15,6] := -0.04656999;
      R_g[15,7] := -0.01576530;
      R_g[15,8] := -0.00584896;
      R_g[15,9] := -0.26015484;
      R_g[15,10] := -0.24142613;
      R_g[15,11] := 0.25730863;
      R_g[15,12] := -0.11453031;
      R_g[15,13] := 0.11119434;
      R_g[15,14] := 0.17737047;
      R_g[15,15] := -2.63738036;
      R_g[15,16] := 0.08244993;
      R_g[15,17] := -0.05181377;
      R_g[15,18] := -0.17019351;
      R_g[15,19] := -0.00057711;
      R_g[15,20] := -0.06410737;
      R_g[15,21] := -0.35635000;
      R_g[15,22] := -0.05634273;
      R_g[15,23] := -0.05787534;
      R_g[15,24] := -0.28821653;
      R_g[15,25] := 0.04072954;
      R_g[15,26] := -0.35264266;
      R_g[15,27] := -0.02693767;
      R_g[15,28] := 0.00252916;
      R_g[15,29] := 0.13764562;
      R_g[15,30] := -0.00824686;
      R_g[15,31] := 0.12128824;
      R_g[16,0] := 0.60132068;
      R_g[16,1] := -0.01856642;
      R_g[16,2] := -0.08966170;
      R_g[16,3] := -0.13946506;
      R_g[16,4] := -0.00415761;
      R_g[16,5] := -0.28280789;
      R_g[16,6] := 0.06967461;
      R_g[16,7] := 0.23631206;
      R_g[16,8] := 0.23964688;
      R_g[16,9] := -0.29860437;
      R_g[16,10] := -0.29331362;
      R_g[16,11] := -0.06584249;
      R_g[16,12] := -0.09147212;
      R_g[16,13] := -0.46546975;
      R_g[16,14] := 0.12629899;
      R_g[16,15] := -0.06389543;
      R_g[16,16] := -0.40778831;
      R_g[16,17] := 0.11143796;
      R_g[16,18] := -0.27378660;
      R_g[16,19] := 0.00952273;
      R_g[16,20] := 0.02246955;
      R_g[16,21] := 0.05861741;
      R_g[16,22] := 0.15492634;
      R_g[16,23] := -0.11301065;
      R_g[16,24] := -0.08985913;
      R_g[16,25] := -0.02188338;
      R_g[16,26] := 0.33387843;
      R_g[16,27] := -0.16640456;
      R_g[16,28] := 0.01505111;
      R_g[16,29] := -0.33711705;
      R_g[16,30] := 0.02125577;
      R_g[16,31] := 0.01524946;
      R_g[17,0] := -0.38925147;
      R_g[17,1] := 0.10167669;
      R_g[17,2] := 1.09963822;
      R_g[17,3] := 0.56638694;
      R_g[17,4] := -0.38925627;
      R_g[17,5] := -0.28342962;
      R_g[17,6] := -0.09601510;
      R_g[17,7] := -0.10801526;
      R_g[17,8] := -0.35662961;
      R_g[17,9] := -0.04573594;
      R_g[17,10] := -0.64441895;
      R_g[17,11] := 0.10761937;
      R_g[17,12] := 0.40848148;
      R_g[17,13] := 0.21693566;
      R_g[17,14] := -0.47779572;
      R_g[17,15] := 0.05735239;
      R_g[17,16] := 0.61725920;
      R_g[17,17] := -0.99182111;
      R_g[17,18] := -0.28720608;
      R_g[17,19] := -0.55444890;
      R_g[17,20] := -0.08293245;
      R_g[17,21] := -0.06818427;
      R_g[17,22] := 0.36398715;
      R_g[17,23] := -0.03210070;
      R_g[17,24] := -0.28585058;
      R_g[17,25] := -0.27513689;
      R_g[17,26] := 0.03552913;
      R_g[17,27] := -0.08013315;
      R_g[17,28] := 0.35897267;
      R_g[17,29] := 0.14637794;
      R_g[17,30] := 0.02656880;
      R_g[17,31] := 0.09042920;
      R_g[18,0] := 0.10600080;
      R_g[18,1] := -0.27434132;
      R_g[18,2] := -0.00969330;
      R_g[18,3] := 0.05851525;
      R_g[18,4] := 0.36833468;
      R_g[18,5] := -0.14349443;
      R_g[18,6] := 0.57578582;
      R_g[18,7] := -0.07903897;
      R_g[18,8] := 0.22599036;
      R_g[18,9] := 0.16850802;
      R_g[18,10] := 0.39619374;
      R_g[18,11] := -0.08689134;
      R_g[18,12] := -0.02203394;
      R_g[18,13] := 0.09214581;
      R_g[18,14] := -0.18136357;
      R_g[18,15] := -0.18521205;
      R_g[18,16] := -0.12584965;
      R_g[18,17] := 0.02805296;
      R_g[18,18] := -2.82306099;
      R_g[18,19] := 0.02860738;
      R_g[18,20] := -0.06768390;
      R_g[18,21] := -0.17756699;
      R_g[18,22] := -0.35438040;
      R_g[18,23] := 0.00587577;
      R_g[18,24] := 0.14259399;
      R_g[18,25] := -0.15871549;
      R_g[18,26] := -0.08291962;
      R_g[18,27] := -0.01776898;
      R_g[18,28] := 0.09889172;
      R_g[18,29] := -0.25204495;
      R_g[18,30] := 0.03351328;
      R_g[18,31] := -0.49044365;
      R_g[19,0] := 0.09904923;
      R_g[19,1] := -0.20450678;
      R_g[19,2] := 0.17437203;
      R_g[19,3] := -0.22587489;
      R_g[19,4] := -0.27591318;
      R_g[19,5] := 0.01043208;
      R_g[19,6] := 0.19569586;
      R_g[19,7] := -0.16759375;
      R_g[19,8] := -0.30989414;
      R_g[19,9] := 0.31677705;
      R_g[19,10] := 0.39843774;
      R_g[19,11] := -0.21896553;
      R_g[19,12] := -0.30846235;
      R_g[19,13] := -0.05650981;
      R_g[19,14] := -0.19992013;
      R_g[19,15] := 0.33444968;
      R_g[19,16] := -0.06378950;
      R_g[19,17] := 0.43867654;
      R_g[19,18] := 0.19880539;
      R_g[19,19] := -0.57955313;
      R_g[19,20] := -0.16816148;
      R_g[19,21] := -0.11770317;
      R_g[19,22] := -0.09540665;
      R_g[19,23] := 0.32714933;
      R_g[19,24] := 0.10426765;
      R_g[19,25] := 0.00905210;
      R_g[19,26] := 0.17375226;
      R_g[19,27] := 0.06059144;
      R_g[19,28] := -0.07685973;
      R_g[19,29] := 0.13111910;
      R_g[19,30] := -0.06328917;
      R_g[19,31] := 0.17372234;
      R_g[20,0] := 0.45158643;
      R_g[20,1] := 0.10048324;
      R_g[20,2] := -0.18336149;
      R_g[20,3] := 0.04757790;
      R_g[20,4] := -0.52304280;
      R_g[20,5] := 0.42825961;
      R_g[20,6] := -0.09577745;
      R_g[20,7] := -0.14495638;
      R_g[20,8] := 0.08802815;
      R_g[20,9] := 0.25205737;
      R_g[20,10] := -0.32155499;
      R_g[20,11] := 0.05428667;
      R_g[20,12] := -0.18616134;
      R_g[20,13] := -0.25662100;
      R_g[20,14] := 0.23557436;
      R_g[20,15] := -0.07531256;
      R_g[20,16] := -0.03767674;
      R_g[20,17] := 0.12337428;
      R_g[20,18] := 0.27934751;
      R_g[20,19] := -0.00926364;
      R_g[20,20] := -3.79986739;
      R_g[20,21] := -0.19543613;
      R_g[20,22] := 0.09970980;
      R_g[20,23] := 0.31888810;
      R_g[20,24] := -0.16263051;
      R_g[20,25] := 0.40389246;
      R_g[20,26] := 0.17506121;
      R_g[20,27] := -0.12197474;
      R_g[20,28] := 0.33344150;
      R_g[20,29] := 0.53447098;
      R_g[20,30] := -0.08177848;
      R_g[20,31] := 0.16116713;
      R_g[21,0] := 0.23435149;
      R_g[21,1] := -0.12724286;
      R_g[21,2] := 0.28686163;
      R_g[21,3] := 0.32758567;
      R_g[21,4] := 0.37008581;
      R_g[21,5] := 0.00054913;
      R_g[21,6] := -0.20666862;
      R_g[21,7] := -0.07006288;
      R_g[21,8] := 0.03611933;
      R_g[21,9] := 0.02129174;
      R_g[21,10] := -0.37161198;
      R_g[21,11] := 0.15757479;
      R_g[21,12] := 0.02570746;
      R_g[21,13] := 0.02327103;
      R_g[21,14] := 0.09640582;
      R_g[21,15] := 0.26042229;
      R_g[21,16] := 0.34472993;
      R_g[21,17] := -0.00835064;
      R_g[21,18] := 0.00551167;
      R_g[21,19] := -0.11429182;
      R_g[21,20] := 0.03507146;
      R_g[21,21] := -3.44825172;
      R_g[21,22] := -0.26649529;
      R_g[21,23] := -0.10135769;
      R_g[21,24] := 0.34481728;
      R_g[21,25] := -0.23443097;
      R_g[21,26] := 0.16992255;
      R_g[21,27] := -0.13308460;
      R_g[21,28] := -0.24103378;
      R_g[21,29] := -0.41093639;
      R_g[21,30] := 0.26364964;
      R_g[21,31] := -0.16022304;
      R_g[22,0] := -0.07493737;
      R_g[22,1] := 0.17759214;
      R_g[22,2] := -0.01062989;
      R_g[22,3] := -0.30531928;
      R_g[22,4] := -0.03052065;
      R_g[22,5] := -0.03414509;
      R_g[22,6] := 0.18659861;
      R_g[22,7] := 0.21062662;
      R_g[22,8] := -0.17346539;
      R_g[22,9] := -0.19939077;
      R_g[22,10] := 0.12670304;
      R_g[22,11] := 0.06660150;
      R_g[22,12] := 0.26966450;
      R_g[22,13] := 0.10541053;
      R_g[22,14] := 0.64287060;
      R_g[22,15] := -0.08089455;
      R_g[22,16] := 0.04482723;
      R_g[22,17] := -0.38308454;
      R_g[22,18] := -0.33886632;
      R_g[22,19] := -0.01181675;
      R_g[22,20] := 0.00163985;
      R_g[22,21] := -0.05718180;
      R_g[22,22] := -3.16081810;
      R_g[22,23] := 0.07466732;
      R_g[22,24] := -0.30864209;
      R_g[22,25] := 0.07774863;
      R_g[22,26] := 0.02183296;
      R_g[22,27] := 0.06526875;
      R_g[22,28] := 0.01511325;
      R_g[22,29] := -0.07152145;
      R_g[22,30] := -0.00525320;
      R_g[22,31] := 0.29649878;
      R_g[23,0] := 0.00113127;
      R_g[23,1] := 0.12522221;
      R_g[23,2] := 0.05907319;
      R_g[23,3] := -0.02262744;
      R_g[23,4] := -0.10188442;
      R_g[23,5] := -0.21190459;
      R_g[23,6] := 0.18007506;
      R_g[23,7] := 0.05896083;
      R_g[23,8] := -0.22042561;
      R_g[23,9] := -0.50632614;
      R_g[23,10] := -0.25184467;
      R_g[23,11] := -0.02071220;
      R_g[23,12] := 0.13488033;
      R_g[23,13] := 0.58272606;
      R_g[23,14] := -0.34117222;
      R_g[23,15] := -0.05228347;
      R_g[23,16] := 0.00460199;
      R_g[23,17] := -0.11781638;
      R_g[23,18] := 0.23311849;
      R_g[23,19] := -0.04014893;
      R_g[23,20] := -0.33957833;
      R_g[23,21] := 0.02890438;
      R_g[23,22] := -0.24083762;
      R_g[23,23] := -0.94268411;
      R_g[23,24] := -0.03553833;
      R_g[23,25] := -0.01412383;
      R_g[23,26] := -0.18156384;
      R_g[23,27] := -0.09131307;
      R_g[23,28] := -0.44586113;
      R_g[23,29] := -0.03801443;
      R_g[23,30] := 0.00086464;
      R_g[23,31] := 0.26916614;
      R_g[24,0] := -0.64336246;
      R_g[24,1] := 0.10306925;
      R_g[24,2] := 0.51399171;
      R_g[24,3] := -0.05540410;
      R_g[24,4] := -0.03185389;
      R_g[24,5] := -0.24791254;
      R_g[24,6] := 0.20463978;
      R_g[24,7] := 0.23886493;
      R_g[24,8] := 0.07842016;
      R_g[24,9] := -0.30920368;
      R_g[24,10] := 0.23489781;
      R_g[24,11] := 0.12703019;
      R_g[24,12] := 0.16607307;
      R_g[24,13] := 0.49904567;
      R_g[24,14] := -0.17724575;
      R_g[24,15] := 0.28705874;
      R_g[24,16] := 0.10735691;
      R_g[24,17] := -0.20810044;
      R_g[24,18] := -0.05945748;
      R_g[24,19] := 0.08566293;
      R_g[24,20] := 0.23888144;
      R_g[24,21] := 0.37153292;
      R_g[24,22] := -0.05995385;
      R_g[24,23] := -0.41755617;
      R_g[24,24] := -3.88887119;
      R_g[24,25] := -0.41723010;
      R_g[24,26] := -0.13346243;
      R_g[24,27] := -0.14061303;
      R_g[24,28] := -0.13331260;
      R_g[24,29] := -0.03063603;
      R_g[24,30] := 0.05910332;
      R_g[24,31] := -0.25991386;
      R_g[25,0] := -0.05274433;
      R_g[25,1] := 0.00594214;
      R_g[25,2] := -0.11314983;
      R_g[25,3] := 0.00570132;
      R_g[25,4] := 0.36403185;
      R_g[25,5] := -0.01250168;
      R_g[25,6] := 0.19910777;
      R_g[25,7] := 0.34642568;
      R_g[25,8] := 0.01872415;
      R_g[25,9] := -0.44597912;
      R_g[25,10] := -0.07655778;
      R_g[25,11] := 0.10288168;
      R_g[25,12] := 0.03142342;
      R_g[25,13] := 0.02222106;
      R_g[25,14] := -0.23081708;
      R_g[25,15] := -0.17446531;
      R_g[25,16] := 0.12313956;
      R_g[25,17] := -0.50936556;
      R_g[25,18] := -0.28882426;
      R_g[25,19] := 0.16454880;
      R_g[25,20] := 0.17461465;
      R_g[25,21] := -0.14967380;
      R_g[25,22] := -0.08211164;
      R_g[25,23] := -0.49162635;
      R_g[25,24] := 0.02804507;
      R_g[25,25] := -3.43903923;
      R_g[25,26] := 0.03487247;
      R_g[25,27] := 0.10763391;
      R_g[25,28] := -0.19208704;
      R_g[25,29] := 0.09429935;
      R_g[25,30] := -0.05688680;
      R_g[25,31] := -0.35967454;
      R_g[26,0] := -0.35371888;
      R_g[26,1] := -0.16951147;
      R_g[26,2] := 0.02608063;
      R_g[26,3] := -0.33375439;
      R_g[26,4] := -0.07263146;
      R_g[26,5] := 0.18195383;
      R_g[26,6] := -0.03087202;
      R_g[26,7] := -0.16634339;
      R_g[26,8] := -0.11040545;
      R_g[26,9] := 0.32063729;
      R_g[26,10] := 0.33352721;
      R_g[26,11] := -0.35319483;
      R_g[26,12] := -0.36759371;
      R_g[26,13] := 0.04302413;
      R_g[26,14] := -0.39809039;
      R_g[26,15] := 0.58213729;
      R_g[26,16] := -0.48063713;
      R_g[26,17] := 0.31698564;
      R_g[26,18] := 0.40641028;
      R_g[26,19] := 0.05107375;
      R_g[26,20] := 0.02146294;
      R_g[26,21] := -0.36092263;
      R_g[26,22] := 0.12869963;
      R_g[26,23] := 0.03362994;
      R_g[26,24] := 0.01885223;
      R_g[26,25] := 0.19347078;
      R_g[26,26] := -3.84916234;
      R_g[26,27] := 0.25620162;
      R_g[26,28] := -0.00354434;
      R_g[26,29] := 0.26753259;
      R_g[26,30] := 0.27058694;
      R_g[26,31] := -0.06458917;
      R_g[27,0] := -0.26864582;
      R_g[27,1] := -0.46819380;
      R_g[27,2] := -0.10896234;
      R_g[27,3] := 0.27843839;
      R_g[27,4] := -0.26515251;
      R_g[27,5] := -0.10256714;
      R_g[27,6] := -0.09258715;
      R_g[27,7] := 0.32607606;
      R_g[27,8] := -0.23709811;
      R_g[27,9] := -0.40867603;
      R_g[27,10] := -0.50749040;
      R_g[27,11] := 0.19362329;
      R_g[27,12] := -0.02271074;
      R_g[27,13] := -0.25827619;
      R_g[27,14] := 0.89860833;
      R_g[27,15] := -0.32963204;
      R_g[27,16] := 0.30623397;
      R_g[27,17] := -0.41240448;
      R_g[27,18] := -0.29421324;
      R_g[27,19] := -0.03716093;
      R_g[27,20] := 0.16659185;
      R_g[27,21] := 0.06818414;
      R_g[27,22] := 0.25484851;
      R_g[27,23] := 0.22020060;
      R_g[27,24] := -0.23671104;
      R_g[27,25] := 0.21126530;
      R_g[27,26] := 0.51748723;
      R_g[27,27] := -3.80495954;
      R_g[27,28] := 0.25846967;
      R_g[27,29] := -0.27945098;
      R_g[27,30] := -0.06130871;
      R_g[27,31] := 0.30456460;
      R_g[28,0] := 0.08912513;
      R_g[28,1] := -0.06453909;
      R_g[28,2] := -0.27234399;
      R_g[28,3] := 0.08671865;
      R_g[28,4] := 0.35958216;
      R_g[28,5] := -0.14240554;
      R_g[28,6] := -0.21201842;
      R_g[28,7] := 0.03412353;
      R_g[28,8] := -0.03125657;
      R_g[28,9] := -0.46181759;
      R_g[28,10] := 0.01940809;
      R_g[28,11] := 0.25482264;
      R_g[28,12] := 0.05732013;
      R_g[28,13] := 0.17726658;
      R_g[28,14] := 0.06626137;
      R_g[28,15] := -0.12480546;
      R_g[28,16] := 0.02746791;
      R_g[28,17] := -0.12780708;
      R_g[28,18] := -0.30959740;
      R_g[28,19] := -0.13992572;
      R_g[28,20] := -0.18084787;
      R_g[28,21] := -0.19184320;
      R_g[28,22] := -0.06709936;
      R_g[28,23] := 0.05110632;
      R_g[28,24] := -0.18117674;
      R_g[28,25] := -0.00072563;
      R_g[28,26] := -0.08458403;
      R_g[28,27] := 0.10861294;
      R_g[28,28] := -2.71115732;
      R_g[28,29] := -0.37569851;
      R_g[28,30] := 0.06543881;
      R_g[28,31] := 0.09642852;
      R_g[29,0] := -0.05788187;
      R_g[29,1] := -0.27650809;
      R_g[29,2] := 0.29699826;
      R_g[29,3] := 0.19907336;
      R_g[29,4] := -0.16655856;
      R_g[29,5] := 0.11022907;
      R_g[29,6] := 0.19868205;
      R_g[29,7] := -0.12020898;
      R_g[29,8] := -0.04434412;
      R_g[29,9] := 0.54825044;
      R_g[29,10] := 0.16285433;
      R_g[29,11] := -0.25309601;
      R_g[29,12] := -0.08369306;
      R_g[29,13] := 0.01308564;
      R_g[29,14] := -0.13750511;
      R_g[29,15] := -0.18384902;
      R_g[29,16] := -0.12176835;
      R_g[29,17] := 0.37266698;
      R_g[29,18] := 0.35773721;
      R_g[29,19] := 0.11458746;
      R_g[29,20] := -0.17479272;
      R_g[29,21] := 0.40825108;
      R_g[29,22] := 0.29202622;
      R_g[29,23] := 0.05949272;
      R_g[29,24] := -0.03869816;
      R_g[29,25] := -0.01413330;
      R_g[29,26] := 0.54103899;
      R_g[29,27] := 0.37894773;
      R_g[29,28] := -0.13715395;
      R_g[29,29] := -2.87533021;
      R_g[29,30] := -0.20007172;
      R_g[29,31] := -0.13430515;
      R_g[30,0] := 0.26030293;
      R_g[30,1] := -0.91468990;
      R_g[30,2] := -0.70711064;
      R_g[30,3] := 0.17348513;
      R_g[30,4] := -0.09719203;
      R_g[30,5] := -0.55125755;
      R_g[30,6] := 0.29799628;
      R_g[30,7] := -0.06895110;
      R_g[30,8] := -0.10511522;
      R_g[30,9] := 0.15847020;
      R_g[30,10] := 0.51417458;
      R_g[30,11] := -0.35962448;
      R_g[30,12] := -0.30896205;
      R_g[30,13] := 0.05734081;
      R_g[30,14] := 0.07842971;
      R_g[30,15] := -0.36382475;
      R_g[30,16] := -0.41747949;
      R_g[30,17] := 0.19075811;
      R_g[30,18] := 0.25313321;
      R_g[30,19] := 0.55022001;
      R_g[30,20] := -0.49628595;
      R_g[30,21] := 0.08953253;
      R_g[30,22] := 0.00409314;
      R_g[30,23] := 0.40932578;
      R_g[30,24] := -0.17622793;
      R_g[30,25] := 0.14825498;
      R_g[30,26] := -0.14895549;
      R_g[30,27] := 0.15221059;
      R_g[30,28] := -0.43621781;
      R_g[30,29] := 1.00098062;
      R_g[30,30] := -2.90753388;
      R_g[30,31] := 0.75884044;
      R_g[31,0] := 0.17272399;
      R_g[31,1] := -0.05801272;
      R_g[31,2] := -0.01508001;
      R_g[31,3] := 0.14520457;
      R_g[31,4] := 0.32392308;
      R_g[31,5] := 0.07295397;
      R_g[31,6] := 0.03031077;
      R_g[31,7] := -0.18328291;
      R_g[31,8] := 0.11090327;
      R_g[31,9] := 0.04064663;
      R_g[31,10] := -0.47682047;
      R_g[31,11] := 0.15038835;
      R_g[31,12] := -0.08792843;
      R_g[31,13] := -0.12402203;
      R_g[31,14] := -0.28880438;
      R_g[31,15] := 0.08178798;
      R_g[31,16] := 0.36903802;
      R_g[31,17] := -0.59405959;
      R_g[31,18] := -0.02349467;
      R_g[31,19] := 0.09523650;
      R_g[31,20] := 0.11543348;
      R_g[31,21] := 0.13315134;
      R_g[31,22] := 0.14046821;
      R_g[31,23] := 0.07318171;
      R_g[31,24] := 0.36266720;
      R_g[31,25] := -0.08543201;
      R_g[31,26] := 0.04509775;
      R_g[31,27] := 0.05353892;
      R_g[31,28] := 0.09169131;
      R_g[31,29] := -0.00655315;
      R_g[31,30] := 0.06718629;
      R_g[31,31] := -2.64188099;
      R_o[0,0] := 2.30278349;
      R_o[0,1] := 0.14783031;
      R_o[0,2] := -4.34446335;
      R_o[0,3] := 0.08713067;
      R_o[0,4] := 0.44618216;
      R_o[0,5] := -0.91748381;
      R_o[0,6] := -0.03610091;
      R_o[0,7] := 0.31388551;
      R_o[0,8] := -0.56839061;
      R_o[0,9] := -1.09572577;
      R_o[0,10] := -0.28296462;
      R_o[0,11] := 0.11638703;
      R_o[0,12] := -0.26847789;
      R_o[0,13] := -2.86956191;
      R_o[0,14] := -0.09927089;
      R_o[0,15] := -0.02761977;
      R_o[0,16] := 0.52737570;
      R_o[0,17] := -0.79886532;
      R_o[0,18] := -0.49760529;
      R_o[0,19] := 0.44731107;
      R_o[0,20] := -0.28426364;
      R_o[0,21] := 0.00891846;
      R_o[0,22] := 0.33747271;
      R_o[0,23] := -0.50627428;
      R_o[0,24] := 2.19249272;
      R_o[0,25] := -0.04657436;
      R_o[0,26] := 0.05185679;
      R_o[0,27] := 0.21695121;
      R_o[0,28] := 0.10701730;
      R_o[0,29] := -0.13881534;
      R_o[0,30] := 0.26203036;
      R_o[0,31] := 0.34208903;
      R_o[1,0] := 0.96568722;
      R_o[1,1] := 3.20853710;
      R_o[1,2] := -0.90170866;
      R_o[1,3] := -0.37756726;
      R_o[1,4] := 0.76046461;
      R_o[1,5] := -1.21417594;
      R_o[1,6] := -0.70202482;
      R_o[1,7] := 0.02065790;
      R_o[1,8] := 0.59182841;
      R_o[1,9] := -0.54165220;
      R_o[1,10] := 0.68561763;
      R_o[1,11] := 0.05523187;
      R_o[1,12] := -0.11933473;
      R_o[1,13] := -0.83110988;
      R_o[1,14] := 0.44425490;
      R_o[1,15] := 0.49311119;
      R_o[1,16] := 0.63592368;
      R_o[1,17] := -0.71622342;
      R_o[1,18] := -0.37737587;
      R_o[1,19] := -0.47871071;
      R_o[1,20] := 0.73954928;
      R_o[1,21] := -0.34349287;
      R_o[1,22] := 0.23899685;
      R_o[1,23] := -0.40250215;
      R_o[1,24] := 0.48065677;
      R_o[1,25] := -0.19839822;
      R_o[1,26] := 0.18214372;
      R_o[1,27] := -0.63379246;
      R_o[1,28] := 1.21917188;
      R_o[1,29] := -0.66983658;
      R_o[1,30] := -0.10998060;
      R_o[1,31] := 0.93811083;
      R_o[2,0] := -0.13516584;
      R_o[2,1] := -0.04461868;
      R_o[2,2] := -0.26925364;
      R_o[2,3] := -0.23952584;
      R_o[2,4] := 0.66424054;
      R_o[2,5] := 0.14358610;
      R_o[2,6] := -0.29987994;
      R_o[2,7] := 0.00934964;
      R_o[2,8] := -0.14183417;
      R_o[2,9] := -0.56005502;
      R_o[2,10] := 0.13025737;
      R_o[2,11] := -0.00965034;
      R_o[2,12] := -0.22625396;
      R_o[2,13] := -1.17763340;
      R_o[2,14] := -0.39688507;
      R_o[2,15] := 0.16797350;
      R_o[2,16] := -0.11934988;
      R_o[2,17] := -0.13632622;
      R_o[2,18] := -0.04847634;
      R_o[2,19] := 0.19914898;
      R_o[2,20] := 0.26995429;
      R_o[2,21] := -0.70818353;
      R_o[2,22] := -0.30348709;
      R_o[2,23] := -0.58659947;
      R_o[2,24] := 1.18079221;
      R_o[2,25] := -0.40847197;
      R_o[2,26] := -0.26015049;
      R_o[2,27] := -1.17746425;
      R_o[2,28] := -0.23879230;
      R_o[2,29] := -0.00942878;
      R_o[2,30] := 0.46976960;
      R_o[2,31] := -0.11859558;
      R_o[3,0] := 0.20476769;
      R_o[3,1] := 0.33900335;
      R_o[3,2] := -0.09836011;
      R_o[3,3] := 1.78037620;
      R_o[3,4] := 0.24503271;
      R_o[3,5] := -0.61845154;
      R_o[3,6] := -0.20356861;
      R_o[3,7] := 0.04746798;
      R_o[3,8] := 0.50998628;
      R_o[3,9] := -0.78148943;
      R_o[3,10] := -0.08412565;
      R_o[3,11] := 0.26778370;
      R_o[3,12] := 0.08690196;
      R_o[3,13] := -0.26804864;
      R_o[3,14] := -0.00070689;
      R_o[3,15] := 0.06325699;
      R_o[3,16] := 0.62193298;
      R_o[3,17] := -0.39169067;
      R_o[3,18] := -0.43697286;
      R_o[3,19] := 0.25084570;
      R_o[3,20] := -0.89430416;
      R_o[3,21] := -0.27173933;
      R_o[3,22] := 1.84822822;
      R_o[3,23] := -0.63409132;
      R_o[3,24] := 1.02836239;
      R_o[3,25] := -0.22855356;
      R_o[3,26] := -0.05025835;
      R_o[3,27] := -0.18045969;
      R_o[3,28] := 0.07945272;
      R_o[3,29] := -0.47019318;
      R_o[3,30] := 0.17809509;
      R_o[3,31] := -0.56552023;
      R_o[4,0] := 0.43562740;
      R_o[4,1] := -0.23176828;
      R_o[4,2] := 0.14830057;
      R_o[4,3] := 0.36350489;
      R_o[4,4] := -0.16774306;
      R_o[4,5] := 0.20693526;
      R_o[4,6] := 0.20155330;
      R_o[4,7] := 0.04864905;
      R_o[4,8] := -0.33429313;
      R_o[4,9] := -0.35912898;
      R_o[4,10] := 0.46565962;
      R_o[4,11] := 0.01946744;
      R_o[4,12] := 0.10726556;
      R_o[4,13] := 0.20833483;
      R_o[4,14] := -0.61803621;
      R_o[4,15] := -0.19495259;
      R_o[4,16] := 0.02558211;
      R_o[4,17] := -0.33150405;
      R_o[4,18] := -0.29833490;
      R_o[4,19] := 0.14919333;
      R_o[4,20] := 0.74265832;
      R_o[4,21] := -0.75234932;
      R_o[4,22] := 0.44413266;
      R_o[4,23] := -0.35464638;
      R_o[4,24] := 0.03076732;
      R_o[4,25] := -0.03035804;
      R_o[4,26] := 0.01813117;
      R_o[4,27] := -0.16126633;
      R_o[4,28] := 0.03274649;
      R_o[4,29] := 0.05024729;
      R_o[4,30] := -0.10365503;
      R_o[4,31] := -0.00369479;
      R_o[5,0] := 0.48018265;
      R_o[5,1] := 0.03282917;
      R_o[5,2] := -0.10870697;
      R_o[5,3] := -0.97790849;
      R_o[5,4] := 0.82862431;
      R_o[5,5] := -1.01685739;
      R_o[5,6] := 0.32942194;
      R_o[5,7] := -0.26762411;
      R_o[5,8] := 0.19432366;
      R_o[5,9] := -0.97326458;
      R_o[5,10] := 0.83567667;
      R_o[5,11] := -0.30151615;
      R_o[5,12] := -0.68087310;
      R_o[5,13] := -1.20724499;
      R_o[5,14] := 0.43663529;
      R_o[5,15] := 0.37139645;
      R_o[5,16] := 0.04509346;
      R_o[5,17] := -0.08997716;
      R_o[5,18] := 0.08793837;
      R_o[5,19] := 0.10307877;
      R_o[5,20] := -0.17214446;
      R_o[5,21] := -0.73129249;
      R_o[5,22] := 1.66565955;
      R_o[5,23] := -0.00417784;
      R_o[5,24] := 0.86307442;
      R_o[5,25] := -0.11585745;
      R_o[5,26] := -0.05403616;
      R_o[5,27] := -0.47711590;
      R_o[5,28] := -0.37349850;
      R_o[5,29] := 1.15859234;
      R_o[5,30] := 0.00607978;
      R_o[5,31] := 0.06847207;
      R_o[6,0] := -0.03867534;
      R_o[6,1] := 0.11462366;
      R_o[6,2] := -0.50761229;
      R_o[6,3] := -0.23780383;
      R_o[6,4] := 0.32394341;
      R_o[6,5] := 0.39529499;
      R_o[6,6] := -0.77105635;
      R_o[6,7] := 0.22093517;
      R_o[6,8] := -0.01466693;
      R_o[6,9] := -0.16930275;
      R_o[6,10] := 0.25404128;
      R_o[6,11] := 0.34278873;
      R_o[6,12] := -0.09828608;
      R_o[6,13] := -0.62504685;
      R_o[6,14] := -0.21883135;
      R_o[6,15] := -0.32010984;
      R_o[6,16] := -0.19807403;
      R_o[6,17] := 0.11536673;
      R_o[6,18] := 0.28473780;
      R_o[6,19] := 0.18543534;
      R_o[6,20] := -0.00624146;
      R_o[6,21] := -0.31709534;
      R_o[6,22] := 0.05469801;
      R_o[6,23] := -0.04293344;
      R_o[6,24] := 0.80048978;
      R_o[6,25] := -0.25435165;
      R_o[6,26] := 0.42625248;
      R_o[6,27] := -0.73878372;
      R_o[6,28] := 0.53613293;
      R_o[6,29] := 0.26586437;
      R_o[6,30] := 0.15208158;
      R_o[6,31] := 0.09870102;
      R_o[7,0] := -0.35428080;
      R_o[7,1] := -0.10483557;
      R_o[7,2] := -0.11971197;
      R_o[7,3] := -0.52425843;
      R_o[7,4] := 0.10465599;
      R_o[7,5] := -0.30066428;
      R_o[7,6] := 0.02017798;
      R_o[7,7] := -0.21352273;
      R_o[7,8] := 0.18289956;
      R_o[7,9] := -0.32229105;
      R_o[7,10] := 0.90695047;
      R_o[7,11] := -0.36772999;
      R_o[7,12] := -0.45428464;
      R_o[7,13] := -0.86696827;
      R_o[7,14] := 0.38000038;
      R_o[7,15] := 0.47287312;
      R_o[7,16] := 0.01553127;
      R_o[7,17] := -0.17758080;
      R_o[7,18] := -0.01059937;
      R_o[7,19] := -0.09118696;
      R_o[7,20] := 0.09259737;
      R_o[7,21] := -0.28630632;
      R_o[7,22] := 0.23516124;
      R_o[7,23] := -0.06806444;
      R_o[7,24] := 0.43746755;
      R_o[7,25] := 0.45478520;
      R_o[7,26] := -0.06099969;
      R_o[7,27] := -0.47780791;
      R_o[7,28] := 0.48667553;
      R_o[7,29] := 0.57442456;
      R_o[7,30] := 0.08897275;
      R_o[7,31] := 0.04724957;
      R_o[8,0] := 0.45044625;
      R_o[8,1] := -0.12919052;
      R_o[8,2] := -0.11546909;
      R_o[8,3] := 0.39766264;
      R_o[8,4] := 0.23777021;
      R_o[8,5] := -0.03082044;
      R_o[8,6] := -0.20632984;
      R_o[8,7] := -0.59559488;
      R_o[8,8] := -0.68259364;
      R_o[8,9] := -0.00083823;
      R_o[8,10] := 0.14988257;
      R_o[8,11] := 0.30479997;
      R_o[8,12] := 0.47008944;
      R_o[8,13] := -0.19031671;
      R_o[8,14] := -0.31048602;
      R_o[8,15] := 0.16468574;
      R_o[8,16] := 0.07428884;
      R_o[8,17] := -0.18089496;
      R_o[8,18] := -0.06553307;
      R_o[8,19] := 0.30119392;
      R_o[8,20] := 0.04313279;
      R_o[8,21] := 0.04614826;
      R_o[8,22] := -0.73448062;
      R_o[8,23] := 0.11781842;
      R_o[8,24] := -0.00477762;
      R_o[8,25] := 0.33527210;
      R_o[8,26] := 0.26166564;
      R_o[8,27] := -0.38534245;
      R_o[8,28] := 0.00645371;
      R_o[8,29] := 0.35132623;
      R_o[8,30] := 0.13199812;
      R_o[8,31] := 0.23807541;
      R_o[9,0] := 0.25993770;
      R_o[9,1] := 0.08555011;
      R_o[9,2] := -0.47537354;
      R_o[9,3] := -0.83094978;
      R_o[9,4] := 0.71708196;
      R_o[9,5] := -0.16037510;
      R_o[9,6] := 0.09589471;
      R_o[9,7] := -0.25086725;
      R_o[9,8] := 0.47328165;
      R_o[9,9] := -0.23029572;
      R_o[9,10] := 0.33668354;
      R_o[9,11] := -0.39398462;
      R_o[9,12] := -0.93957061;
      R_o[9,13] := -0.35627630;
      R_o[9,14] := -0.96541286;
      R_o[9,15] := 0.27267876;
      R_o[9,16] := 0.21410845;
      R_o[9,17] := -0.65840012;
      R_o[9,18] := 0.15242729;
      R_o[9,19] := -0.03121080;
      R_o[9,20] := -0.11927066;
      R_o[9,21] := 0.52784294;
      R_o[9,22] := 0.04285750;
      R_o[9,23] := 0.13811226;
      R_o[9,24] := 0.22844416;
      R_o[9,25] := 0.23292424;
      R_o[9,26] := 0.52570170;
      R_o[9,27] := 0.07966270;
      R_o[9,28] := -0.32864538;
      R_o[9,29] := -0.16931652;
      R_o[9,30] := -0.01193482;
      R_o[9,31] := 0.25869036;
      R_o[10,0] := 0.89997160;
      R_o[10,1] := 0.52300185;
      R_o[10,2] := -0.36115131;
      R_o[10,3] := -0.50931239;
      R_o[10,4] := 0.01933937;
      R_o[10,5] := -0.66100568;
      R_o[10,6] := -0.72948444;
      R_o[10,7] := -0.38120693;
      R_o[10,8] := 0.52716947;
      R_o[10,9] := -0.78645134;
      R_o[10,10] := -0.97260189;
      R_o[10,11] := 0.20774882;
      R_o[10,12] := -0.35503402;
      R_o[10,13] := -0.00724730;
      R_o[10,14] := -1.14668894;
      R_o[10,15] := -0.00573723;
      R_o[10,16] := 0.45797586;
      R_o[10,17] := -0.16783185;
      R_o[10,18] := -0.78439027;
      R_o[10,19] := -0.07787321;
      R_o[10,20] := -0.27455541;
      R_o[10,21] := -0.38741615;
      R_o[10,22] := 2.45607543;
      R_o[10,23] := -0.41554567;
      R_o[10,24] := 0.81808698;
      R_o[10,25] := 0.66784626;
      R_o[10,26] := 0.25790057;
      R_o[10,27] := 0.64080191;
      R_o[10,28] := 0.05862263;
      R_o[10,29] := -0.86733270;
      R_o[10,30] := 0.28249276;
      R_o[10,31] := 0.66749090;
      R_o[11,0] := 0.45413589;
      R_o[11,1] := 0.38346776;
      R_o[11,2] := -0.85281456;
      R_o[11,3] := -0.19667329;
      R_o[11,4] := 0.49708343;
      R_o[11,5] := -0.22616820;
      R_o[11,6] := -0.22052550;
      R_o[11,7] := -0.14427526;
      R_o[11,8] := 0.62248898;
      R_o[11,9] := -1.07283175;
      R_o[11,10] := 0.99012190;
      R_o[11,11] := -0.00387567;
      R_o[11,12] := -0.03953788;
      R_o[11,13] := -0.11381141;
      R_o[11,14] := -0.50175935;
      R_o[11,15] := 0.81905180;
      R_o[11,16] := 0.26642680;
      R_o[11,17] := -0.64103836;
      R_o[11,18] := -0.37297282;
      R_o[11,19] := 0.38684547;
      R_o[11,20] := -0.10901120;
      R_o[11,21] := -0.79144758;
      R_o[11,22] := 0.30630803;
      R_o[11,23] := -0.46943784;
      R_o[11,24] := -0.03455164;
      R_o[11,25] := 0.10039959;
      R_o[11,26] := -0.68668705;
      R_o[11,27] := -0.12410130;
      R_o[11,28] := -0.56831688;
      R_o[11,29] := -0.19138084;
      R_o[11,30] := 0.32598269;
      R_o[11,31] := 0.24842253;
      R_o[12,0] := 0.79577845;
      R_o[12,1] := 1.12471819;
      R_o[12,2] := 0.21189122;
      R_o[12,3] := 0.60872358;
      R_o[12,4] := 0.12913147;
      R_o[12,5] := -0.23679182;
      R_o[12,6] := 0.56693274;
      R_o[12,7] := 0.21713342;
      R_o[12,8] := 0.75730407;
      R_o[12,9] := -1.11194956;
      R_o[12,10] := -0.05170097;
      R_o[12,11] := -0.13823876;
      R_o[12,12] := 2.48078752;
      R_o[12,13] := -0.40249935;
      R_o[12,14] := 0.31937549;
      R_o[12,15] := 0.79539752;
      R_o[12,16] := 1.96585226;
      R_o[12,17] := -0.21539992;
      R_o[12,18] := -0.28552079;
      R_o[12,19] := -0.31043211;
      R_o[12,20] := -0.31463060;
      R_o[12,21] := -0.09506584;
      R_o[12,22] := 1.57885945;
      R_o[12,23] := -0.32251796;
      R_o[12,24] := 0.74886376;
      R_o[12,25] := -0.00495276;
      R_o[12,26] := 0.03871931;
      R_o[12,27] := 0.03866331;
      R_o[12,28] := 0.72467947;
      R_o[12,29] := -0.63773739;
      R_o[12,30] := 0.09163156;
      R_o[12,31] := 0.24973899;
      R_o[13,0] := -0.04444838;
      R_o[13,1] := -0.03776657;
      R_o[13,2] := -1.29966748;
      R_o[13,3] := -1.21049142;
      R_o[13,4] := 0.61895919;
      R_o[13,5] := 0.42413464;
      R_o[13,6] := -0.26110905;
      R_o[13,7] := 0.01253382;
      R_o[13,8] := 0.67533016;
      R_o[13,9] := -1.22368360;
      R_o[13,10] := 1.24057198;
      R_o[13,11] := -0.26758894;
      R_o[13,12] := 0.06042844;
      R_o[13,13] := -0.04051395;
      R_o[13,14] := 1.54065347;
      R_o[13,15] := 1.18497789;
      R_o[13,16] := 0.45765820;
      R_o[13,17] := -0.53086120;
      R_o[13,18] := 0.18301466;
      R_o[13,19] := 0.70264763;
      R_o[13,20] := 0.52861190;
      R_o[13,21] := -1.26863003;
      R_o[13,22] := 0.67413718;
      R_o[13,23] := -0.77813780;
      R_o[13,24] := 2.00173545;
      R_o[13,25] := -0.20376748;
      R_o[13,26] := -0.36850744;
      R_o[13,27] := -1.54971695;
      R_o[13,28] := -0.18608753;
      R_o[13,29] := 0.25340420;
      R_o[13,30] := 0.79221284;
      R_o[13,31] := -0.22243516;
      R_o[14,0] := 0.36772186;
      R_o[14,1] := 0.35438997;
      R_o[14,2] := 0.79816318;
      R_o[14,3] := -0.71921414;
      R_o[14,4] := 0.01499140;
      R_o[14,5] := -0.16665320;
      R_o[14,6] := 0.54814249;
      R_o[14,7] := -0.31334832;
      R_o[14,8] := 1.54228234;
      R_o[14,9] := -0.38194096;
      R_o[14,10] := -0.16915111;
      R_o[14,11] := -0.35635409;
      R_o[14,12] := -0.09595951;
      R_o[14,13] := 1.54526842;
      R_o[14,14] := 3.68650222;
      R_o[14,15] := 0.04523968;
      R_o[14,16] := 0.68481857;
      R_o[14,17] := -0.30135879;
      R_o[14,18] := 0.04055335;
      R_o[14,19] := 0.19981964;
      R_o[14,20] := -1.15916789;
      R_o[14,21] := -0.61886412;
      R_o[14,22] := 2.11957574;
      R_o[14,23] := -0.04530338;
      R_o[14,24] := 0.23210397;
      R_o[14,25] := 0.34942800;
      R_o[14,26] := 0.39147028;
      R_o[14,27] := 0.58273619;
      R_o[14,28] := -1.05760503;
      R_o[14,29] := 0.24741873;
      R_o[14,30] := 0.16608724;
      R_o[14,31] := 0.39260611;
      R_o[15,0] := 0.51947361;
      R_o[15,1] := -0.12846206;
      R_o[15,2] := -0.66827095;
      R_o[15,3] := 0.56208074;
      R_o[15,4] := 0.22565739;
      R_o[15,5] := -0.55710828;
      R_o[15,6] := -0.64466113;
      R_o[15,7] := 0.36292467;
      R_o[15,8] := 0.50899130;
      R_o[15,9] := -0.74116105;
      R_o[15,10] := 0.08156371;
      R_o[15,11] := 0.57796168;
      R_o[15,12] := -0.26711142;
      R_o[15,13] := 0.71900034;
      R_o[15,14] := 0.45004350;
      R_o[15,15] := -2.02677822;
      R_o[15,16] := 0.17003906;
      R_o[15,17] := -0.78767359;
      R_o[15,18] := -0.42787877;
      R_o[15,19] := -0.36432889;
      R_o[15,20] := -0.36618990;
      R_o[15,21] := -0.97692233;
      R_o[15,22] := 0.27408621;
      R_o[15,23] := -0.24445024;
      R_o[15,24] := 0.07183556;
      R_o[15,25] := -0.13564034;
      R_o[15,26] := -0.20052052;
      R_o[15,27] := 0.06819152;
      R_o[15,28] := 0.00067334;
      R_o[15,29] := -0.31617504;
      R_o[15,30] := -0.25879920;
      R_o[15,31] := 0.59753007;
      R_o[16,0] := 0.28681985;
      R_o[16,1] := -0.34336987;
      R_o[16,2] := 0.50298339;
      R_o[16,3] := -0.43604618;
      R_o[16,4] := 0.19562161;
      R_o[16,5] := -0.54955274;
      R_o[16,6] := -0.02381020;
      R_o[16,7] := 0.34711182;
      R_o[16,8] := 0.89456636;
      R_o[16,9] := -0.28739411;
      R_o[16,10] := 0.36038986;
      R_o[16,11] := 0.34008405;
      R_o[16,12] := -0.37093174;
      R_o[16,13] := 0.36884668;
      R_o[16,14] := -0.10169870;
      R_o[16,15] := -0.47918934;
      R_o[16,16] := 1.61680961;
      R_o[16,17] := -0.97384298;
      R_o[16,18] := -0.04127910;
      R_o[16,19] := -0.22060362;
      R_o[16,20] := -0.02375492;
      R_o[16,21] := 0.09434792;
      R_o[16,22] := 0.43916631;
      R_o[16,23] := -0.49490130;
      R_o[16,24] := 0.34134132;
      R_o[16,25] := -0.54296613;
      R_o[16,26] := -0.01715025;
      R_o[16,27] := -0.37928930;
      R_o[16,28] := -0.19477750;
      R_o[16,29] := 0.24976863;
      R_o[16,30] := -0.11030178;
      R_o[16,31] := -0.19956882;
      R_o[17,0] := 0.48948678;
      R_o[17,1] := -0.00858265;
      R_o[17,2] := -0.24564666;
      R_o[17,3] := -0.15596397;
      R_o[17,4] := 0.46464425;
      R_o[17,5] := -0.52813530;
      R_o[17,6] := 0.47345904;
      R_o[17,7] := 0.01340096;
      R_o[17,8] := -0.26542130;
      R_o[17,9] := -0.11717621;
      R_o[17,10] := 0.54016209;
      R_o[17,11] := 0.20284952;
      R_o[17,12] := 0.02328762;
      R_o[17,13] := 0.12176004;
      R_o[17,14] := -0.58269668;
      R_o[17,15] := 0.07123553;
      R_o[17,16] := -0.39322037;
      R_o[17,17] := -0.10467571;
      R_o[17,18] := -0.06699307;
      R_o[17,19] := 0.31953976;
      R_o[17,20] := -0.28262883;
      R_o[17,21] := -0.12952352;
      R_o[17,22] := 0.12820345;
      R_o[17,23] := -0.59919792;
      R_o[17,24] := 0.25555119;
      R_o[17,25] := -0.05377883;
      R_o[17,26] := -0.00513316;
      R_o[17,27] := 0.07034966;
      R_o[17,28] := 0.16618735;
      R_o[17,29] := 0.12366936;
      R_o[17,30] := 0.11204547;
      R_o[17,31] := -0.36965579;
      R_o[18,0] := 0.28828311;
      R_o[18,1] := -0.00360730;
      R_o[18,2] := -0.66725665;
      R_o[18,3] := -0.44986060;
      R_o[18,4] := -0.15414765;
      R_o[18,5] := -0.68566316;
      R_o[18,6] := 0.33631477;
      R_o[18,7] := -0.56416988;
      R_o[18,8] := -0.32173297;
      R_o[18,9] := -0.16714011;
      R_o[18,10] := 0.13619064;
      R_o[18,11] := -0.35170969;
      R_o[18,12] := -0.51983321;
      R_o[18,13] := 0.21738678;
      R_o[18,14] := -0.08145608;
      R_o[18,15] := 0.01709783;
      R_o[18,16] := -0.18718076;
      R_o[18,17] := -0.40229329;
      R_o[18,18] := -0.24698442;
      R_o[18,19] := -0.23457956;
      R_o[18,20] := -0.39634994;
      R_o[18,21] := -0.06818978;
      R_o[18,22] := -0.37303329;
      R_o[18,23] := 0.00050139;
      R_o[18,24] := 0.67526346;
      R_o[18,25] := 0.45440361;
      R_o[18,26] := 0.69033909;
      R_o[18,27] := -0.46217164;
      R_o[18,28] := 0.14283627;
      R_o[18,29] := -0.15705536;
      R_o[18,30] := 0.21938857;
      R_o[18,31] := 0.46284494;
      R_o[19,0] := 0.97230667;
      R_o[19,1] := 0.96507812;
      R_o[19,2] := -0.57360196;
      R_o[19,3] := -1.02491653;
      R_o[19,4] := 1.00897348;
      R_o[19,5] := -0.00255713;
      R_o[19,6] := -0.35491705;
      R_o[19,7] := -0.29408309;
      R_o[19,8] := -0.29375651;
      R_o[19,9] := -0.46368971;
      R_o[19,10] := 0.73696595;
      R_o[19,11] := 0.09828018;
      R_o[19,12] := 0.55897504;
      R_o[19,13] := -0.14518775;
      R_o[19,14] := -0.04863453;
      R_o[19,15] := 1.61602235;
      R_o[19,16] := 0.05364607;
      R_o[19,17] := -0.13429411;
      R_o[19,18] := -0.06690535;
      R_o[19,19] := 0.08334047;
      R_o[19,20] := 0.13419743;
      R_o[19,21] := -0.19960804;
      R_o[19,22] := 1.20868075;
      R_o[19,23] := -0.96787804;
      R_o[19,24] := 0.87696582;
      R_o[19,25] := -0.06458701;
      R_o[19,26] := 0.28224054;
      R_o[19,27] := -0.96385705;
      R_o[19,28] := -0.54325783;
      R_o[19,29] := -1.00623095;
      R_o[19,30] := 0.23156840;
      R_o[19,31] := 0.29148033;
      R_o[20,0] := -0.15315647;
      R_o[20,1] := -0.09547617;
      R_o[20,2] := -0.46687099;
      R_o[20,3] := 0.11482628;
      R_o[20,4] := 0.67318785;
      R_o[20,5] := 0.15630811;
      R_o[20,6] := -0.43997395;
      R_o[20,7] := 0.21123159;
      R_o[20,8] := -0.04171057;
      R_o[20,9] := -0.65907657;
      R_o[20,10] := 0.42881182;
      R_o[20,11] := 0.07429390;
      R_o[20,12] := -0.50155687;
      R_o[20,13] := -0.66903663;
      R_o[20,14] := -0.32008776;
      R_o[20,15] := -0.22985753;
      R_o[20,16] := 0.05104850;
      R_o[20,17] := -0.36443755;
      R_o[20,18] := -0.04919767;
      R_o[20,19] := 0.10203130;
      R_o[20,20] := -0.11491112;
      R_o[20,21] := -0.70318282;
      R_o[20,22] := -0.08754787;
      R_o[20,23] := -0.47064683;
      R_o[20,24] := 0.23331608;
      R_o[20,25] := -0.03932161;
      R_o[20,26] := -0.05192051;
      R_o[20,27] := -0.40804467;
      R_o[20,28] := 0.16400859;
      R_o[20,29] := -0.02629855;
      R_o[20,30] := 0.34915683;
      R_o[20,31] := -0.04184714;
      R_o[21,0] := 0.66911119;
      R_o[21,1] := 0.00413969;
      R_o[21,2] := -0.20499986;
      R_o[21,3] := -0.68706846;
      R_o[21,4] := 0.43500739;
      R_o[21,5] := -0.77048969;
      R_o[21,6] := 0.43577152;
      R_o[21,7] := -0.41412577;
      R_o[21,8] := -0.23024948;
      R_o[21,9] := -0.14370334;
      R_o[21,10] := 0.19276123;
      R_o[21,11] := -0.45450440;
      R_o[21,12] := -0.17385210;
      R_o[21,13] := -0.43938136;
      R_o[21,14] := -0.15357804;
      R_o[21,15] := -0.36838773;
      R_o[21,16] := 0.12680964;
      R_o[21,17] := -0.72252679;
      R_o[21,18] := -0.17201090;
      R_o[21,19] := -0.75203276;
      R_o[21,20] := 0.45121738;
      R_o[21,21] := 2.52927732;
      R_o[21,22] := 2.61969614;
      R_o[21,23] := -0.12567814;
      R_o[21,24] := 0.33255699;
      R_o[21,25] := 0.49635842;
      R_o[21,26] := 0.89324474;
      R_o[21,27] := -1.15636325;
      R_o[21,28] := 1.21784663;
      R_o[21,29] := -0.30604303;
      R_o[21,30] := -0.73844993;
      R_o[21,31] := -0.77427286;
      R_o[22,0] := 0.26138592;
      R_o[22,1] := 0.04288378;
      R_o[22,2] := -0.23030537;
      R_o[22,3] := 0.07515529;
      R_o[22,4] := 0.17849518;
      R_o[22,5] := -0.22360083;
      R_o[22,6] := -0.99275935;
      R_o[22,7] := -0.25043544;
      R_o[22,8] := 0.16721144;
      R_o[22,9] := -0.59967136;
      R_o[22,10] := 0.40209976;
      R_o[22,11] := 0.16054669;
      R_o[22,12] := -0.13949765;
      R_o[22,13] := -0.73240519;
      R_o[22,14] := -0.22012003;
      R_o[22,15] := 0.01868595;
      R_o[22,16] := 0.34183541;
      R_o[22,17] := 0.02852705;
      R_o[22,18] := -0.04114153;
      R_o[22,19] := -0.00736952;
      R_o[22,20] := -0.15057497;
      R_o[22,21] := -0.41413474;
      R_o[22,22] := 0.76486248;
      R_o[22,23] := -0.76816767;
      R_o[22,24] := 0.05123224;
      R_o[22,25] := 0.13371366;
      R_o[22,26] := 0.05483653;
      R_o[22,27] := 0.43419600;
      R_o[22,28] := -0.05295467;
      R_o[22,29] := -0.13698067;
      R_o[22,30] := -0.27184281;
      R_o[22,31] := 0.68283230;
      R_o[23,0] := 0.15452501;
      R_o[23,1] := 0.38931781;
      R_o[23,2] := -0.71978974;
      R_o[23,3] := -0.11382619;
      R_o[23,4] := 0.32177678;
      R_o[23,5] := 0.53753215;
      R_o[23,6] := 0.10605058;
      R_o[23,7] := 0.15947971;
      R_o[23,8] := 0.05374712;
      R_o[23,9] := -0.03133825;
      R_o[23,10] := 0.12940039;
      R_o[23,11] := -0.58461565;
      R_o[23,12] := -0.24854553;
      R_o[23,13] := -0.37112287;
      R_o[23,14] := 0.04672547;
      R_o[23,15] := -0.00671248;
      R_o[23,16] := -0.09047767;
      R_o[23,17] := -0.83457744;
      R_o[23,18] := -0.47293767;
      R_o[23,19] := -0.31071156;
      R_o[23,20] := 0.03737261;
      R_o[23,21] := -0.31324276;
      R_o[23,22] := -0.01070617;
      R_o[23,23] := 1.53010750;
      R_o[23,24] := 0.23675759;
      R_o[23,25] := 0.10948038;
      R_o[23,26] := 0.46215081;
      R_o[23,27] := -0.36760142;
      R_o[23,28] := 0.75483471;
      R_o[23,29] := -0.15528834;
      R_o[23,30] := 0.01413946;
      R_o[23,31] := -0.38331240;
      R_o[24,0] := -0.10675674;
      R_o[24,1] := -0.51453239;
      R_o[24,2] := -0.00356475;
      R_o[24,3] := -0.16368514;
      R_o[24,4] := 0.13058373;
      R_o[24,5] := 0.37898996;
      R_o[24,6] := -0.04559740;
      R_o[24,7] := 0.32021171;
      R_o[24,8] := 0.87053347;
      R_o[24,9] := -0.38837278;
      R_o[24,10] := 0.52733487;
      R_o[24,11] := 0.13364539;
      R_o[24,12] := -0.66372377;
      R_o[24,13] := -0.32406506;
      R_o[24,14] := 0.58510506;
      R_o[24,15] := 0.16703159;
      R_o[24,16] := -0.03636205;
      R_o[24,17] := -0.74969834;
      R_o[24,18] := 0.04493890;
      R_o[24,19] := 0.07232044;
      R_o[24,20] := -0.72455716;
      R_o[24,21] := -0.71928841;
      R_o[24,22] := 1.00345361;
      R_o[24,23] := -0.10275900;
      R_o[24,24] := 0.14540374;
      R_o[24,25] := 0.08173257;
      R_o[24,26] := 0.01965822;
      R_o[24,27] := -0.48747879;
      R_o[24,28] := 0.38453004;
      R_o[24,29] := 0.15411790;
      R_o[24,30] := 0.12267981;
      R_o[24,31] := -0.25638211;
      R_o[25,0] := 0.50944263;
      R_o[25,1] := -0.10795844;
      R_o[25,2] := -0.69347328;
      R_o[25,3] := -0.57176161;
      R_o[25,4] := 0.86021614;
      R_o[25,5] := 0.17890315;
      R_o[25,6] := -0.49303707;
      R_o[25,7] := 0.42926988;
      R_o[25,8] := 0.03010171;
      R_o[25,9] := -0.46701196;
      R_o[25,10] := 0.22579275;
      R_o[25,11] := 0.00480429;
      R_o[25,12] := 0.11027759;
      R_o[25,13] := -0.36264303;
      R_o[25,14] := 0.11242234;
      R_o[25,15] := 0.17056607;
      R_o[25,16] := -0.01122399;
      R_o[25,17] := -0.50582260;
      R_o[25,18] := -0.55902225;
      R_o[25,19] := 0.05534580;
      R_o[25,20] := -0.34148753;
      R_o[25,21] := -0.14953679;
      R_o[25,22] := -0.16325586;
      R_o[25,23] := 0.00732038;
      R_o[25,24] := -0.03740266;
      R_o[25,25] := -0.32909846;
      R_o[25,26] := -0.10309041;
      R_o[25,27] := -0.22430740;
      R_o[25,28] := 0.16309188;
      R_o[25,29] := 0.32213110;
      R_o[25,30] := 0.18461545;
      R_o[25,31] := -0.05051695;
      R_o[26,0] := 0.49827960;
      R_o[26,1] := 0.28162920;
      R_o[26,2] := -2.07256627;
      R_o[26,3] := -0.71399188;
      R_o[26,4] := 0.15465102;
      R_o[26,5] := 0.02878987;
      R_o[26,6] := -0.59221852;
      R_o[26,7] := -0.38292849;
      R_o[26,8] := 1.90265203;
      R_o[26,9] := -0.72589833;
      R_o[26,10] := -0.03948683;
      R_o[26,11] := -0.33430120;
      R_o[26,12] := -0.78429389;
      R_o[26,13] := 0.00490210;
      R_o[26,14] := -0.73278040;
      R_o[26,15] := 0.19303162;
      R_o[26,16] := 0.65501148;
      R_o[26,17] := -0.87329102;
      R_o[26,18] := 0.02019684;
      R_o[26,19] := -0.33091050;
      R_o[26,20] := -0.27779147;
      R_o[26,21] := -2.15610600;
      R_o[26,22] := -0.04925109;
      R_o[26,23] := -0.50757724;
      R_o[26,24] := -0.06259642;
      R_o[26,25] := -0.11439695;
      R_o[26,26] := -3.03007960;
      R_o[26,27] := -0.26429990;
      R_o[26,28] := 0.24497572;
      R_o[26,29] := 0.23329099;
      R_o[26,30] := 0.65626943;
      R_o[26,31] := 0.82046634;
      R_o[27,0] := -0.25980654;
      R_o[27,1] := -0.85493249;
      R_o[27,2] := -0.25568795;
      R_o[27,3] := -0.11439860;
      R_o[27,4] := 0.10520780;
      R_o[27,5] := -0.15565851;
      R_o[27,6] := 0.01195115;
      R_o[27,7] := -0.07017966;
      R_o[27,8] := -0.03355999;
      R_o[27,9] := -0.21074077;
      R_o[27,10] := 0.03461521;
      R_o[27,11] := 0.07374318;
      R_o[27,12] := -0.22766791;
      R_o[27,13] := -0.78329474;
      R_o[27,14] := -0.30588287;
      R_o[27,15] := 0.71185470;
      R_o[27,16] := -0.11062124;
      R_o[27,17] := 0.15082856;
      R_o[27,18] := -0.00008092;
      R_o[27,19] := 0.06574772;
      R_o[27,20] := 0.39814237;
      R_o[27,21] := 0.41286281;
      R_o[27,22] := -0.35842898;
      R_o[27,23] := -0.14691216;
      R_o[27,24] := 0.45409301;
      R_o[27,25] := 0.06740260;
      R_o[27,26] := 0.18736783;
      R_o[27,27] := -0.82008070;
      R_o[27,28] := -0.21420176;
      R_o[27,29] := 0.49815652;
      R_o[27,30] := 0.13462545;
      R_o[27,31] := -0.44356906;
      R_o[28,0] := 0.41890109;
      R_o[28,1] := 0.01776026;
      R_o[28,2] := -0.60563636;
      R_o[28,3] := -0.60062194;
      R_o[28,4] := 0.60836959;
      R_o[28,5] := -0.00771509;
      R_o[28,6] := -0.38145909;
      R_o[28,7] := 0.40494025;
      R_o[28,8] := -0.34993392;
      R_o[28,9] := 0.00921785;
      R_o[28,10] := -0.08201695;
      R_o[28,11] := 0.21442677;
      R_o[28,12] := 0.01693209;
      R_o[28,13] := -0.03023057;
      R_o[28,14] := -0.71048105;
      R_o[28,15] := 0.13766295;
      R_o[28,16] := -0.06296610;
      R_o[28,17] := -0.30172476;
      R_o[28,18] := -0.31208399;
      R_o[28,19] := 0.52773523;
      R_o[28,20] := 0.44576228;
      R_o[28,21] := -0.62207425;
      R_o[28,22] := 0.49633217;
      R_o[28,23] := 0.00518359;
      R_o[28,24] := 0.42131236;
      R_o[28,25] := -0.34798115;
      R_o[28,26] := -0.02231124;
      R_o[28,27] := -0.29808775;
      R_o[28,28] := 0.54361582;
      R_o[28,29] := 0.29003334;
      R_o[28,30] := 0.40789396;
      R_o[28,31] := -0.06554151;
      R_o[29,0] := 0.02121896;
      R_o[29,1] := 0.09064472;
      R_o[29,2] := 0.31729925;
      R_o[29,3] := 0.10008687;
      R_o[29,4] := 0.17747171;
      R_o[29,5] := -0.11045200;
      R_o[29,6] := 0.11371059;
      R_o[29,7] := -0.23605901;
      R_o[29,8] := -0.08776284;
      R_o[29,9] := 0.32796374;
      R_o[29,10] := 0.15019821;
      R_o[29,11] := -0.22550444;
      R_o[29,12] := -0.01797267;
      R_o[29,13] := -0.35675609;
      R_o[29,14] := -0.74846828;
      R_o[29,15] := 0.04661415;
      R_o[29,16] := -0.06017135;
      R_o[29,17] := -0.03003342;
      R_o[29,18] := 0.24155578;
      R_o[29,19] := 0.09004185;
      R_o[29,20] := -0.14736657;
      R_o[29,21] := -0.14575130;
      R_o[29,22] := 0.12607163;
      R_o[29,23] := -0.22345687;
      R_o[29,24] := 0.15827295;
      R_o[29,25] := 0.02486655;
      R_o[29,26] := -0.10162737;
      R_o[29,27] := -0.17148840;
      R_o[29,28] := -0.04898299;
      R_o[29,29] := 0.96720076;
      R_o[29,30] := -0.07629140;
      R_o[29,31] := -0.11269102;
      R_o[30,0] := -0.33895251;
      R_o[30,1] := -0.45090100;
      R_o[30,2] := -0.63235575;
      R_o[30,3] := -0.11448206;
      R_o[30,4] := 0.44136623;
      R_o[30,5] := -0.15951085;
      R_o[30,6] := -0.19755951;
      R_o[30,7] := 0.09543595;
      R_o[30,8] := 0.50030470;
      R_o[30,9] := 0.25317916;
      R_o[30,10] := 0.21241242;
      R_o[30,11] := -0.12849870;
      R_o[30,12] := -0.63707429;
      R_o[30,13] := -0.03736546;
      R_o[30,14] := -0.47734249;
      R_o[30,15] := -1.42653191;
      R_o[30,16] := -0.49558908;
      R_o[30,17] := -0.00803843;
      R_o[30,18] := 0.10319717;
      R_o[30,19] := 0.01286428;
      R_o[30,20] := 0.16171345;
      R_o[30,21] := -0.07717690;
      R_o[30,22] := -0.23527963;
      R_o[30,23] := 0.55368316;
      R_o[30,24] := 0.90191066;
      R_o[30,25] := -0.44086981;
      R_o[30,26] := -0.32070184;
      R_o[30,27] := -0.45357138;
      R_o[30,28] := 0.02687183;
      R_o[30,29] := 0.03311172;
      R_o[30,30] := -1.04822719;
      R_o[30,31] := 0.29971805;
      R_o[31,0] := 0.12431819;
      R_o[31,1] := 0.23183918;
      R_o[31,2] := -0.30574140;
      R_o[31,3] := -0.59901828;
      R_o[31,4] := 0.05242074;
      R_o[31,5] := 0.22697972;
      R_o[31,6] := -0.01884122;
      R_o[31,7] := -0.17017308;
      R_o[31,8] := 0.33408687;
      R_o[31,9] := -0.04179906;
      R_o[31,10] := -0.12077110;
      R_o[31,11] := 0.28922603;
      R_o[31,12] := -0.08880246;
      R_o[31,13] := -0.15585485;
      R_o[31,14] := -0.02141503;
      R_o[31,15] := 0.21018416;
      R_o[31,16] := -0.09174474;
      R_o[31,17] := -0.46324244;
      R_o[31,18] := -0.46089089;
      R_o[31,19] := -0.02686797;
      R_o[31,20] := 0.07938531;
      R_o[31,21] := -0.19916745;
      R_o[31,22] := -0.38484034;
      R_o[31,23] := -0.01166240;
      R_o[31,24] := 0.13159335;
      R_o[31,25] := 0.12521118;
      R_o[31,26] := 0.03883914;
      R_o[31,27] := 0.04080096;
      R_o[31,28] := -0.01131530;
      R_o[31,29] := -0.18011786;
      R_o[31,30] := 0.12775224;
      R_o[31,31] := 0.56156427;
      B_i[0] := -0.11037196;
      B_i[1] := -0.20119080;
      B_i[2] := -0.47118652;
      B_i[3] := -0.26821959;
      B_i[4] := -0.06291195;
      B_i[5] := -0.34240282;
      B_i[6] := 0.06325857;
      B_i[7] := 0.45427629;
      B_i[8] := 0.66686732;
      B_i[9] := 0.18742950;
      B_i[10] := -0.70640790;
      B_i[11] := 0.02270032;
      B_i[12] := 0.22158253;
      B_i[13] := -1.29529023;
      B_i[14] := -0.54597330;
      B_i[15] := -0.11060837;
      B_i[16] := 1.80296397;
      B_i[17] := -0.12063497;
      B_i[18] := 0.05746642;
      B_i[19] := 0.38928580;
      B_i[20] := -0.31188878;
      B_i[21] := -0.24247971;
      B_i[22] := -0.31664434;
      B_i[23] := 1.62169862;
      B_i[24] := -0.90392292;
      B_i[25] := -0.15748771;
      B_i[26] := 0.13672107;
      B_i[27] := -0.39835182;
      B_i[28] := -0.01372162;
      B_i[29] := 2.23123884;
      B_i[30] := 1.44870400;
      B_i[31] := 0.68679756;
      B_f[0] := 4.12368870;
      B_f[1] := 2.80252981;
      B_f[2] := 3.82664418;
      B_f[3] := -1.81176567;
      B_f[4] := -0.07009026;
      B_f[5] := 3.66103506;
      B_f[6] := 2.19355917;
      B_f[7] := 1.98418212;
      B_f[8] := -1.10244370;
      B_f[9] := -1.93180275;
      B_f[10] := -4.32190752;
      B_f[11] := 1.51885438;
      B_f[12] := 1.65448213;
      B_f[13] := 4.53528595;
      B_f[14] := -0.56549478;
      B_f[15] := 0.10521974;
      B_f[16] := -1.76427710;
      B_f[17] := -0.08624527;
      B_f[18] := 3.21538043;
      B_f[19] := -1.63178980;
      B_f[20] := 3.08151102;
      B_f[21] := 1.74406099;
      B_f[22] := 1.94425082;
      B_f[23] := -0.94436306;
      B_f[24] := 2.89898777;
      B_f[25] := 2.95786500;
      B_f[26] := 1.61822867;
      B_f[27] := 2.82563996;
      B_f[28] := 2.15152121;
      B_f[29] := 3.32113457;
      B_f[30] := -0.17399743;
      B_f[31] := 0.91838026;
      B_g[0] := 0.95918286;
      B_g[1] := 0.20353325;
      B_g[2] := -0.46430916;
      B_g[3] := -1.68014383;
      B_g[4] := 0.58820122;
      B_g[5] := 0.03108167;
      B_g[6] := -0.24217492;
      B_g[7] := -0.00992692;
      B_g[8] := 0.45266634;
      B_g[9] := -1.96682358;
      B_g[10] := 0.25125173;
      B_g[11] := 0.32966834;
      B_g[12] := 0.22510809;
      B_g[13] := -0.84138256;
      B_g[14] := 0.85291719;
      B_g[15] := -0.23710170;
      B_g[16] := 0.40418231;
      B_g[17] := -1.26592064;
      B_g[18] := 0.32817277;
      B_g[19] := 0.36937705;
      B_g[20] := 0.07663520;
      B_g[21] := 0.08663416;
      B_g[22] := 0.47949010;
      B_g[23] := -0.28541470;
      B_g[24] := 0.76597357;
      B_g[25] := 0.03829502;
      B_g[26] := 0.86952877;
      B_g[27] := -0.31516683;
      B_g[28] := -0.22333460;
      B_g[29] := -0.05720093;
      B_g[30] := 0.66168761;
      B_g[31] := -0.39613989;
      B_o[0] := 2.81217766;
      B_o[1] := 3.59746456;
      B_o[2] := 2.71275401;
      B_o[3] := 1.75578141;
      B_o[4] := 0.73969102;
      B_o[5] := 3.72038746;
      B_o[6] := 1.89435756;
      B_o[7] := 3.43835115;
      B_o[8] := 1.45377648;
      B_o[9] := 3.22759438;
      B_o[10] := 2.52799082;
      B_o[11] := 3.16732812;
      B_o[12] := 3.56140375;
      B_o[13] := 4.45837831;
      B_o[14] := 3.20861292;
      B_o[15] := -0.15407386;
      B_o[16] := 2.85862112;
      B_o[17] := 1.02626765;
      B_o[18] := 3.48203158;
      B_o[19] := 3.79925871;
      B_o[20] := 1.95770288;
      B_o[21] := 2.69921970;
      B_o[22] := 2.34376049;
      B_o[23] := 1.60421276;
      B_o[24] := 2.49631310;
      B_o[25] := 2.75451827;
      B_o[26] := 3.84688234;
      B_o[27] := 2.41971064;
      B_o[28] := 2.71536970;
      B_o[29] := 0.46796203;
      B_o[30] := 1.03240466;
      B_o[31] := 2.02655077;
      FC_W[0,0] := -0.91911894;
      FC_W[0,1] := 1.92505515;
      FC_W[0,2] := -0.46473372;
      FC_W[0,3] := 0.49914464;
      FC_W[0,4] := -0.22144756;
      FC_W[0,5] := -0.10570145;
      FC_W[0,6] := -0.53842652;
      FC_W[0,7] := -0.56898397;
      FC_W[0,8] := 0.62797409;
      FC_W[0,9] := 0.89987290;
      FC_W[0,10] := 0.06315278;
      FC_W[0,11] := 0.68087977;
      FC_W[0,12] := -1.31657398;
      FC_W[0,13] := 0.19018160;
      FC_W[0,14] := 0.30356276;
      FC_W[0,15] := -0.00683733;
      FC_W[0,16] := 0.03132518;
      FC_W[0,17] := -0.47817189;
      FC_W[0,18] := -1.06647837;
      FC_W[0,19] := 0.18862465;
      FC_W[0,20] := -0.26146525;
      FC_W[0,21] := 0.00500324;
      FC_W[0,22] := 0.35247201;
      FC_W[0,23] := -0.11869892;
      FC_W[0,24] := -0.02369487;
      FC_W[0,25] := 0.21972799;
      FC_W[0,26] := 0.27597019;
      FC_W[0,27] := -0.92189664;
      FC_W[0,28] := -0.66625625;
      FC_W[0,29] := 0.11222937;
      FC_W[0,30] := 0.08014797;
      FC_W[0,31] := 0.23311555;
      FC_W[1,0] := 2.24038744;
      FC_W[1,1] := 0.43658215;
      FC_W[1,2] := -0.03753655;
      FC_W[1,3] := 0.28978097;
      FC_W[1,4] := -0.44472128;
      FC_W[1,5] := 2.58052659;
      FC_W[1,6] := 0.22744730;
      FC_W[1,7] := 0.19882494;
      FC_W[1,8] := -0.21679716;
